BEGIN
   Id := 5;
   CancelOrders := FALSE;
   PauseOrders := FALSE;
   ResumeOrders := FALSE;
   OrderSent := FALSE;
   CurrentOrder := 0;
   NextOrder := 1;
   OrderTable[0].OrderNo := 0;
   OrderTable[0].StepNo := 256;
   OrderTable[0].PlaceTime := '';
   OrderTable[0].Device := '';
   OrderTable[0].Sequence := 0;
   OrderTable[0].Status := 'Error';
   OrderTable[0].CompleteTime := '06/10/2022 08:58:15';
   OrderTable[0].ErrorID := 0;
   OrderTable[1].OrderNo := 0;
   OrderTable[1].StepNo := 0;
   OrderTable[1].PlaceTime := '';
   OrderTable[1].Device := '';
   OrderTable[1].Sequence := 0;
   OrderTable[1].Status := '';
   OrderTable[1].CompleteTime := '';
   OrderTable[1].ErrorID := 0;
   OrderTable[2].OrderNo := 0;
   OrderTable[2].StepNo := 0;
   OrderTable[2].PlaceTime := '';
   OrderTable[2].Device := '';
   OrderTable[2].Sequence := 0;
   OrderTable[2].Status := '';
   OrderTable[2].CompleteTime := '';
   OrderTable[2].ErrorID := 0;
   OrderTable[3].OrderNo := 0;
   OrderTable[3].StepNo := 0;
   OrderTable[3].PlaceTime := '';
   OrderTable[3].Device := '';
   OrderTable[3].Sequence := 0;
   OrderTable[3].Status := '';
   OrderTable[3].CompleteTime := '';
   OrderTable[3].ErrorID := 0;
   OrderTable[4].OrderNo := 0;
   OrderTable[4].StepNo := 0;
   OrderTable[4].PlaceTime := '';
   OrderTable[4].Device := '';
   OrderTable[4].Sequence := 0;
   OrderTable[4].Status := '';
   OrderTable[4].CompleteTime := '';
   OrderTable[4].ErrorID := 0;
   OrderTable[5].OrderNo := 0;
   OrderTable[5].StepNo := 0;
   OrderTable[5].PlaceTime := '';
   OrderTable[5].Device := '';
   OrderTable[5].Sequence := 0;
   OrderTable[5].Status := '';
   OrderTable[5].CompleteTime := '';
   OrderTable[5].ErrorID := 0;
   OrderTable[6].OrderNo := 0;
   OrderTable[6].StepNo := 0;
   OrderTable[6].PlaceTime := '';
   OrderTable[6].Device := '';
   OrderTable[6].Sequence := 0;
   OrderTable[6].Status := '';
   OrderTable[6].CompleteTime := '';
   OrderTable[6].ErrorID := 0;
   OrderTable[7].OrderNo := 0;
   OrderTable[7].StepNo := 0;
   OrderTable[7].PlaceTime := '';
   OrderTable[7].Device := '';
   OrderTable[7].Sequence := 0;
   OrderTable[7].Status := '';
   OrderTable[7].CompleteTime := '';
   OrderTable[7].ErrorID := 0;
   OrderTable[8].OrderNo := 0;
   OrderTable[8].StepNo := 0;
   OrderTable[8].PlaceTime := '';
   OrderTable[8].Device := '';
   OrderTable[8].Sequence := 0;
   OrderTable[8].Status := '';
   OrderTable[8].CompleteTime := '';
   OrderTable[8].ErrorID := 0;
   OrderTable[9].OrderNo := 0;
   OrderTable[9].StepNo := 0;
   OrderTable[9].PlaceTime := '';
   OrderTable[9].Device := '';
   OrderTable[9].Sequence := 0;
   OrderTable[9].Status := '';
   OrderTable[9].CompleteTime := '';
   OrderTable[9].ErrorID := 0;
   OrderTable[10].OrderNo := 0;
   OrderTable[10].StepNo := 0;
   OrderTable[10].PlaceTime := '';
   OrderTable[10].Device := '';
   OrderTable[10].Sequence := 0;
   OrderTable[10].Status := '';
   OrderTable[10].CompleteTime := '';
   OrderTable[10].ErrorID := 0;
   OrderTable[11].OrderNo := 0;
   OrderTable[11].StepNo := 0;
   OrderTable[11].PlaceTime := '';
   OrderTable[11].Device := '';
   OrderTable[11].Sequence := 0;
   OrderTable[11].Status := '';
   OrderTable[11].CompleteTime := '';
   OrderTable[11].ErrorID := 0;
   OrderTable[12].OrderNo := 0;
   OrderTable[12].StepNo := 0;
   OrderTable[12].PlaceTime := '';
   OrderTable[12].Device := '';
   OrderTable[12].Sequence := 0;
   OrderTable[12].Status := '';
   OrderTable[12].CompleteTime := '';
   OrderTable[12].ErrorID := 0;
   OrderTable[13].OrderNo := 0;
   OrderTable[13].StepNo := 0;
   OrderTable[13].PlaceTime := '';
   OrderTable[13].Device := '';
   OrderTable[13].Sequence := 0;
   OrderTable[13].Status := '';
   OrderTable[13].CompleteTime := '';
   OrderTable[13].ErrorID := 0;
   OrderTable[14].OrderNo := 0;
   OrderTable[14].StepNo := 0;
   OrderTable[14].PlaceTime := '';
   OrderTable[14].Device := '';
   OrderTable[14].Sequence := 0;
   OrderTable[14].Status := '';
   OrderTable[14].CompleteTime := '';
   OrderTable[14].ErrorID := 0;
   OrderTable[15].OrderNo := 0;
   OrderTable[15].StepNo := 0;
   OrderTable[15].PlaceTime := '';
   OrderTable[15].Device := '';
   OrderTable[15].Sequence := 0;
   OrderTable[15].Status := '';
   OrderTable[15].CompleteTime := '';
   OrderTable[15].ErrorID := 0;
   OrderTable[16].OrderNo := 0;
   OrderTable[16].StepNo := 0;
   OrderTable[16].PlaceTime := '';
   OrderTable[16].Device := '';
   OrderTable[16].Sequence := 0;
   OrderTable[16].Status := '';
   OrderTable[16].CompleteTime := '';
   OrderTable[16].ErrorID := 0;
   OrderTable[17].OrderNo := 0;
   OrderTable[17].StepNo := 0;
   OrderTable[17].PlaceTime := '';
   OrderTable[17].Device := '';
   OrderTable[17].Sequence := 0;
   OrderTable[17].Status := '';
   OrderTable[17].CompleteTime := '';
   OrderTable[17].ErrorID := 0;
   OrderTable[18].OrderNo := 0;
   OrderTable[18].StepNo := 0;
   OrderTable[18].PlaceTime := '';
   OrderTable[18].Device := '';
   OrderTable[18].Sequence := 0;
   OrderTable[18].Status := '';
   OrderTable[18].CompleteTime := '';
   OrderTable[18].ErrorID := 0;
   OrderTable[19].OrderNo := 0;
   OrderTable[19].StepNo := 0;
   OrderTable[19].PlaceTime := '';
   OrderTable[19].Device := '';
   OrderTable[19].Sequence := 0;
   OrderTable[19].Status := '';
   OrderTable[19].CompleteTime := '';
   OrderTable[19].ErrorID := 0;
   OrderTable[20].OrderNo := 0;
   OrderTable[20].StepNo := 0;
   OrderTable[20].PlaceTime := '';
   OrderTable[20].Device := '';
   OrderTable[20].Sequence := 0;
   OrderTable[20].Status := '';
   OrderTable[20].CompleteTime := '';
   OrderTable[20].ErrorID := 0;
   OrderTable[21].OrderNo := 0;
   OrderTable[21].StepNo := 0;
   OrderTable[21].PlaceTime := '';
   OrderTable[21].Device := '';
   OrderTable[21].Sequence := 0;
   OrderTable[21].Status := '';
   OrderTable[21].CompleteTime := '';
   OrderTable[21].ErrorID := 0;
   OrderTable[22].OrderNo := 0;
   OrderTable[22].StepNo := 0;
   OrderTable[22].PlaceTime := '';
   OrderTable[22].Device := '';
   OrderTable[22].Sequence := 0;
   OrderTable[22].Status := '';
   OrderTable[22].CompleteTime := '';
   OrderTable[22].ErrorID := 0;
   OrderTable[23].OrderNo := 0;
   OrderTable[23].StepNo := 0;
   OrderTable[23].PlaceTime := '';
   OrderTable[23].Device := '';
   OrderTable[23].Sequence := 0;
   OrderTable[23].Status := '';
   OrderTable[23].CompleteTime := '';
   OrderTable[23].ErrorID := 0;
   OrderTable[24].OrderNo := 0;
   OrderTable[24].StepNo := 0;
   OrderTable[24].PlaceTime := '';
   OrderTable[24].Device := '';
   OrderTable[24].Sequence := 0;
   OrderTable[24].Status := '';
   OrderTable[24].CompleteTime := '';
   OrderTable[24].ErrorID := 0;
   OrderTable[25].OrderNo := 0;
   OrderTable[25].StepNo := 0;
   OrderTable[25].PlaceTime := '';
   OrderTable[25].Device := '';
   OrderTable[25].Sequence := 0;
   OrderTable[25].Status := '';
   OrderTable[25].CompleteTime := '';
   OrderTable[25].ErrorID := 0;
   OrderTable[26].OrderNo := 0;
   OrderTable[26].StepNo := 0;
   OrderTable[26].PlaceTime := '';
   OrderTable[26].Device := '';
   OrderTable[26].Sequence := 0;
   OrderTable[26].Status := '';
   OrderTable[26].CompleteTime := '';
   OrderTable[26].ErrorID := 0;
   OrderTable[27].OrderNo := 0;
   OrderTable[27].StepNo := 0;
   OrderTable[27].PlaceTime := '';
   OrderTable[27].Device := '';
   OrderTable[27].Sequence := 0;
   OrderTable[27].Status := '';
   OrderTable[27].CompleteTime := '';
   OrderTable[27].ErrorID := 0;
   OrderTable[28].OrderNo := 0;
   OrderTable[28].StepNo := 0;
   OrderTable[28].PlaceTime := '';
   OrderTable[28].Device := '';
   OrderTable[28].Sequence := 0;
   OrderTable[28].Status := '';
   OrderTable[28].CompleteTime := '';
   OrderTable[28].ErrorID := 0;
   OrderTable[29].OrderNo := 0;
   OrderTable[29].StepNo := 0;
   OrderTable[29].PlaceTime := '';
   OrderTable[29].Device := '';
   OrderTable[29].Sequence := 0;
   OrderTable[29].Status := '';
   OrderTable[29].CompleteTime := '';
   OrderTable[29].ErrorID := 0;
   OrderTable[30].OrderNo := 0;
   OrderTable[30].StepNo := 0;
   OrderTable[30].PlaceTime := '';
   OrderTable[30].Device := '';
   OrderTable[30].Sequence := 0;
   OrderTable[30].Status := '';
   OrderTable[30].CompleteTime := '';
   OrderTable[30].ErrorID := 0;
   OrderTable[31].OrderNo := 0;
   OrderTable[31].StepNo := 0;
   OrderTable[31].PlaceTime := '';
   OrderTable[31].Device := '';
   OrderTable[31].Sequence := 0;
   OrderTable[31].Status := '';
   OrderTable[31].CompleteTime := '';
   OrderTable[31].ErrorID := 0;
   OrderTable[32].OrderNo := 0;
   OrderTable[32].StepNo := 0;
   OrderTable[32].PlaceTime := '';
   OrderTable[32].Device := '';
   OrderTable[32].Sequence := 0;
   OrderTable[32].Status := '';
   OrderTable[32].CompleteTime := '';
   OrderTable[32].ErrorID := 0;
   OrderTable[33].OrderNo := 0;
   OrderTable[33].StepNo := 0;
   OrderTable[33].PlaceTime := '';
   OrderTable[33].Device := '';
   OrderTable[33].Sequence := 0;
   OrderTable[33].Status := '';
   OrderTable[33].CompleteTime := '';
   OrderTable[33].ErrorID := 0;
   OrderTable[34].OrderNo := 0;
   OrderTable[34].StepNo := 0;
   OrderTable[34].PlaceTime := '';
   OrderTable[34].Device := '';
   OrderTable[34].Sequence := 0;
   OrderTable[34].Status := '';
   OrderTable[34].CompleteTime := '';
   OrderTable[34].ErrorID := 0;
   OrderTable[35].OrderNo := 0;
   OrderTable[35].StepNo := 0;
   OrderTable[35].PlaceTime := '';
   OrderTable[35].Device := '';
   OrderTable[35].Sequence := 0;
   OrderTable[35].Status := '';
   OrderTable[35].CompleteTime := '';
   OrderTable[35].ErrorID := 0;
   OrderTable[36].OrderNo := 0;
   OrderTable[36].StepNo := 0;
   OrderTable[36].PlaceTime := '';
   OrderTable[36].Device := '';
   OrderTable[36].Sequence := 0;
   OrderTable[36].Status := '';
   OrderTable[36].CompleteTime := '';
   OrderTable[36].ErrorID := 0;
   OrderTable[37].OrderNo := 0;
   OrderTable[37].StepNo := 0;
   OrderTable[37].PlaceTime := '';
   OrderTable[37].Device := '';
   OrderTable[37].Sequence := 0;
   OrderTable[37].Status := '';
   OrderTable[37].CompleteTime := '';
   OrderTable[37].ErrorID := 0;
   OrderTable[38].OrderNo := 0;
   OrderTable[38].StepNo := 0;
   OrderTable[38].PlaceTime := '';
   OrderTable[38].Device := '';
   OrderTable[38].Sequence := 0;
   OrderTable[38].Status := '';
   OrderTable[38].CompleteTime := '';
   OrderTable[38].ErrorID := 0;
   OrderTable[39].OrderNo := 0;
   OrderTable[39].StepNo := 0;
   OrderTable[39].PlaceTime := '';
   OrderTable[39].Device := '';
   OrderTable[39].Sequence := 0;
   OrderTable[39].Status := '';
   OrderTable[39].CompleteTime := '';
   OrderTable[39].ErrorID := 0;
   OrderTable[40].OrderNo := 0;
   OrderTable[40].StepNo := 0;
   OrderTable[40].PlaceTime := '';
   OrderTable[40].Device := '';
   OrderTable[40].Sequence := 0;
   OrderTable[40].Status := '';
   OrderTable[40].CompleteTime := '';
   OrderTable[40].ErrorID := 0;
   OrderTable[41].OrderNo := 0;
   OrderTable[41].StepNo := 0;
   OrderTable[41].PlaceTime := '';
   OrderTable[41].Device := '';
   OrderTable[41].Sequence := 0;
   OrderTable[41].Status := '';
   OrderTable[41].CompleteTime := '';
   OrderTable[41].ErrorID := 0;
   OrderTable[42].OrderNo := 0;
   OrderTable[42].StepNo := 0;
   OrderTable[42].PlaceTime := '';
   OrderTable[42].Device := '';
   OrderTable[42].Sequence := 0;
   OrderTable[42].Status := '';
   OrderTable[42].CompleteTime := '';
   OrderTable[42].ErrorID := 0;
   OrderTable[43].OrderNo := 0;
   OrderTable[43].StepNo := 0;
   OrderTable[43].PlaceTime := '';
   OrderTable[43].Device := '';
   OrderTable[43].Sequence := 0;
   OrderTable[43].Status := '';
   OrderTable[43].CompleteTime := '';
   OrderTable[43].ErrorID := 0;
   OrderTable[44].OrderNo := 0;
   OrderTable[44].StepNo := 0;
   OrderTable[44].PlaceTime := '';
   OrderTable[44].Device := '';
   OrderTable[44].Sequence := 0;
   OrderTable[44].Status := '';
   OrderTable[44].CompleteTime := '';
   OrderTable[44].ErrorID := 0;
   OrderTable[45].OrderNo := 0;
   OrderTable[45].StepNo := 0;
   OrderTable[45].PlaceTime := '';
   OrderTable[45].Device := '';
   OrderTable[45].Sequence := 0;
   OrderTable[45].Status := '';
   OrderTable[45].CompleteTime := '';
   OrderTable[45].ErrorID := 0;
   OrderTable[46].OrderNo := 0;
   OrderTable[46].StepNo := 0;
   OrderTable[46].PlaceTime := '';
   OrderTable[46].Device := '';
   OrderTable[46].Sequence := 0;
   OrderTable[46].Status := '';
   OrderTable[46].CompleteTime := '';
   OrderTable[46].ErrorID := 0;
   OrderTable[47].OrderNo := 0;
   OrderTable[47].StepNo := 0;
   OrderTable[47].PlaceTime := '';
   OrderTable[47].Device := '';
   OrderTable[47].Sequence := 0;
   OrderTable[47].Status := '';
   OrderTable[47].CompleteTime := '';
   OrderTable[47].ErrorID := 0;
   OrderTable[48].OrderNo := 0;
   OrderTable[48].StepNo := 0;
   OrderTable[48].PlaceTime := '';
   OrderTable[48].Device := '';
   OrderTable[48].Sequence := 0;
   OrderTable[48].Status := '';
   OrderTable[48].CompleteTime := '';
   OrderTable[48].ErrorID := 0;
   OrderTable[49].OrderNo := 0;
   OrderTable[49].StepNo := 0;
   OrderTable[49].PlaceTime := '';
   OrderTable[49].Device := '';
   OrderTable[49].Sequence := 0;
   OrderTable[49].Status := '';
   OrderTable[49].CompleteTime := '';
   OrderTable[49].ErrorID := 0;
   OrderTable[50].OrderNo := 0;
   OrderTable[50].StepNo := 0;
   OrderTable[50].PlaceTime := '';
   OrderTable[50].Device := '';
   OrderTable[50].Sequence := 0;
   OrderTable[50].Status := '';
   OrderTable[50].CompleteTime := '';
   OrderTable[50].ErrorID := 0;
   OrderTable[51].OrderNo := 0;
   OrderTable[51].StepNo := 0;
   OrderTable[51].PlaceTime := '';
   OrderTable[51].Device := '';
   OrderTable[51].Sequence := 0;
   OrderTable[51].Status := '';
   OrderTable[51].CompleteTime := '';
   OrderTable[51].ErrorID := 0;
   OrderTable[52].OrderNo := 0;
   OrderTable[52].StepNo := 0;
   OrderTable[52].PlaceTime := '';
   OrderTable[52].Device := '';
   OrderTable[52].Sequence := 0;
   OrderTable[52].Status := '';
   OrderTable[52].CompleteTime := '';
   OrderTable[52].ErrorID := 0;
   OrderTable[53].OrderNo := 0;
   OrderTable[53].StepNo := 0;
   OrderTable[53].PlaceTime := '';
   OrderTable[53].Device := '';
   OrderTable[53].Sequence := 0;
   OrderTable[53].Status := '';
   OrderTable[53].CompleteTime := '';
   OrderTable[53].ErrorID := 0;
   OrderTable[54].OrderNo := 0;
   OrderTable[54].StepNo := 0;
   OrderTable[54].PlaceTime := '';
   OrderTable[54].Device := '';
   OrderTable[54].Sequence := 0;
   OrderTable[54].Status := '';
   OrderTable[54].CompleteTime := '';
   OrderTable[54].ErrorID := 0;
   OrderTable[55].OrderNo := 0;
   OrderTable[55].StepNo := 0;
   OrderTable[55].PlaceTime := '';
   OrderTable[55].Device := '';
   OrderTable[55].Sequence := 0;
   OrderTable[55].Status := '';
   OrderTable[55].CompleteTime := '';
   OrderTable[55].ErrorID := 0;
   OrderTable[56].OrderNo := 0;
   OrderTable[56].StepNo := 0;
   OrderTable[56].PlaceTime := '';
   OrderTable[56].Device := '';
   OrderTable[56].Sequence := 0;
   OrderTable[56].Status := '';
   OrderTable[56].CompleteTime := '';
   OrderTable[56].ErrorID := 0;
   OrderTable[57].OrderNo := 0;
   OrderTable[57].StepNo := 0;
   OrderTable[57].PlaceTime := '';
   OrderTable[57].Device := '';
   OrderTable[57].Sequence := 0;
   OrderTable[57].Status := '';
   OrderTable[57].CompleteTime := '';
   OrderTable[57].ErrorID := 0;
   OrderTable[58].OrderNo := 0;
   OrderTable[58].StepNo := 0;
   OrderTable[58].PlaceTime := '';
   OrderTable[58].Device := '';
   OrderTable[58].Sequence := 0;
   OrderTable[58].Status := '';
   OrderTable[58].CompleteTime := '';
   OrderTable[58].ErrorID := 0;
   OrderTable[59].OrderNo := 0;
   OrderTable[59].StepNo := 0;
   OrderTable[59].PlaceTime := '';
   OrderTable[59].Device := '';
   OrderTable[59].Sequence := 0;
   OrderTable[59].Status := '';
   OrderTable[59].CompleteTime := '';
   OrderTable[59].ErrorID := 0;
   OrderTable[60].OrderNo := 0;
   OrderTable[60].StepNo := 0;
   OrderTable[60].PlaceTime := '';
   OrderTable[60].Device := '';
   OrderTable[60].Sequence := 0;
   OrderTable[60].Status := '';
   OrderTable[60].CompleteTime := '';
   OrderTable[60].ErrorID := 0;
   OrderTable[61].OrderNo := 0;
   OrderTable[61].StepNo := 0;
   OrderTable[61].PlaceTime := '';
   OrderTable[61].Device := '';
   OrderTable[61].Sequence := 0;
   OrderTable[61].Status := '';
   OrderTable[61].CompleteTime := '';
   OrderTable[61].ErrorID := 0;
   OrderTable[62].OrderNo := 0;
   OrderTable[62].StepNo := 0;
   OrderTable[62].PlaceTime := '';
   OrderTable[62].Device := '';
   OrderTable[62].Sequence := 0;
   OrderTable[62].Status := '';
   OrderTable[62].CompleteTime := '';
   OrderTable[62].ErrorID := 0;
   OrderTable[63].OrderNo := 0;
   OrderTable[63].StepNo := 0;
   OrderTable[63].PlaceTime := '';
   OrderTable[63].Device := '';
   OrderTable[63].Sequence := 0;
   OrderTable[63].Status := '';
   OrderTable[63].CompleteTime := '';
   OrderTable[63].ErrorID := 0;
   OrderTable[64].OrderNo := 0;
   OrderTable[64].StepNo := 0;
   OrderTable[64].PlaceTime := '';
   OrderTable[64].Device := '';
   OrderTable[64].Sequence := 0;
   OrderTable[64].Status := '';
   OrderTable[64].CompleteTime := '';
   OrderTable[64].ErrorID := 0;
   OrderTable[65].OrderNo := 0;
   OrderTable[65].StepNo := 0;
   OrderTable[65].PlaceTime := '';
   OrderTable[65].Device := '';
   OrderTable[65].Sequence := 0;
   OrderTable[65].Status := '';
   OrderTable[65].CompleteTime := '';
   OrderTable[65].ErrorID := 0;
   OrderTable[66].OrderNo := 0;
   OrderTable[66].StepNo := 0;
   OrderTable[66].PlaceTime := '';
   OrderTable[66].Device := '';
   OrderTable[66].Sequence := 0;
   OrderTable[66].Status := '';
   OrderTable[66].CompleteTime := '';
   OrderTable[66].ErrorID := 0;
   OrderTable[67].OrderNo := 0;
   OrderTable[67].StepNo := 0;
   OrderTable[67].PlaceTime := '';
   OrderTable[67].Device := '';
   OrderTable[67].Sequence := 0;
   OrderTable[67].Status := '';
   OrderTable[67].CompleteTime := '';
   OrderTable[67].ErrorID := 0;
   OrderTable[68].OrderNo := 0;
   OrderTable[68].StepNo := 0;
   OrderTable[68].PlaceTime := '';
   OrderTable[68].Device := '';
   OrderTable[68].Sequence := 0;
   OrderTable[68].Status := '';
   OrderTable[68].CompleteTime := '';
   OrderTable[68].ErrorID := 0;
   OrderTable[69].OrderNo := 0;
   OrderTable[69].StepNo := 0;
   OrderTable[69].PlaceTime := '';
   OrderTable[69].Device := '';
   OrderTable[69].Sequence := 0;
   OrderTable[69].Status := '';
   OrderTable[69].CompleteTime := '';
   OrderTable[69].ErrorID := 0;
   OrderTable[70].OrderNo := 0;
   OrderTable[70].StepNo := 0;
   OrderTable[70].PlaceTime := '';
   OrderTable[70].Device := '';
   OrderTable[70].Sequence := 0;
   OrderTable[70].Status := '';
   OrderTable[70].CompleteTime := '';
   OrderTable[70].ErrorID := 0;
   OrderTable[71].OrderNo := 0;
   OrderTable[71].StepNo := 0;
   OrderTable[71].PlaceTime := '';
   OrderTable[71].Device := '';
   OrderTable[71].Sequence := 0;
   OrderTable[71].Status := '';
   OrderTable[71].CompleteTime := '';
   OrderTable[71].ErrorID := 0;
   OrderTable[72].OrderNo := 0;
   OrderTable[72].StepNo := 0;
   OrderTable[72].PlaceTime := '';
   OrderTable[72].Device := '';
   OrderTable[72].Sequence := 0;
   OrderTable[72].Status := '';
   OrderTable[72].CompleteTime := '';
   OrderTable[72].ErrorID := 0;
   OrderTable[73].OrderNo := 0;
   OrderTable[73].StepNo := 0;
   OrderTable[73].PlaceTime := '';
   OrderTable[73].Device := '';
   OrderTable[73].Sequence := 0;
   OrderTable[73].Status := '';
   OrderTable[73].CompleteTime := '';
   OrderTable[73].ErrorID := 0;
   OrderTable[74].OrderNo := 0;
   OrderTable[74].StepNo := 0;
   OrderTable[74].PlaceTime := '';
   OrderTable[74].Device := '';
   OrderTable[74].Sequence := 0;
   OrderTable[74].Status := '';
   OrderTable[74].CompleteTime := '';
   OrderTable[74].ErrorID := 0;
   OrderTable[75].OrderNo := 0;
   OrderTable[75].StepNo := 0;
   OrderTable[75].PlaceTime := '';
   OrderTable[75].Device := '';
   OrderTable[75].Sequence := 0;
   OrderTable[75].Status := '';
   OrderTable[75].CompleteTime := '';
   OrderTable[75].ErrorID := 0;
   OrderTable[76].OrderNo := 0;
   OrderTable[76].StepNo := 0;
   OrderTable[76].PlaceTime := '';
   OrderTable[76].Device := '';
   OrderTable[76].Sequence := 0;
   OrderTable[76].Status := '';
   OrderTable[76].CompleteTime := '';
   OrderTable[76].ErrorID := 0;
   OrderTable[77].OrderNo := 0;
   OrderTable[77].StepNo := 0;
   OrderTable[77].PlaceTime := '';
   OrderTable[77].Device := '';
   OrderTable[77].Sequence := 0;
   OrderTable[77].Status := '';
   OrderTable[77].CompleteTime := '';
   OrderTable[77].ErrorID := 0;
   OrderTable[78].OrderNo := 0;
   OrderTable[78].StepNo := 0;
   OrderTable[78].PlaceTime := '';
   OrderTable[78].Device := '';
   OrderTable[78].Sequence := 0;
   OrderTable[78].Status := '';
   OrderTable[78].CompleteTime := '';
   OrderTable[78].ErrorID := 0;
   OrderTable[79].OrderNo := 0;
   OrderTable[79].StepNo := 0;
   OrderTable[79].PlaceTime := '';
   OrderTable[79].Device := '';
   OrderTable[79].Sequence := 0;
   OrderTable[79].Status := '';
   OrderTable[79].CompleteTime := '';
   OrderTable[79].ErrorID := 0;
   OrderTable[80].OrderNo := 0;
   OrderTable[80].StepNo := 0;
   OrderTable[80].PlaceTime := '';
   OrderTable[80].Device := '';
   OrderTable[80].Sequence := 0;
   OrderTable[80].Status := '';
   OrderTable[80].CompleteTime := '';
   OrderTable[80].ErrorID := 0;
   OrderTable[81].OrderNo := 0;
   OrderTable[81].StepNo := 0;
   OrderTable[81].PlaceTime := '';
   OrderTable[81].Device := '';
   OrderTable[81].Sequence := 0;
   OrderTable[81].Status := '';
   OrderTable[81].CompleteTime := '';
   OrderTable[81].ErrorID := 0;
   OrderTable[82].OrderNo := 0;
   OrderTable[82].StepNo := 0;
   OrderTable[82].PlaceTime := '';
   OrderTable[82].Device := '';
   OrderTable[82].Sequence := 0;
   OrderTable[82].Status := '';
   OrderTable[82].CompleteTime := '';
   OrderTable[82].ErrorID := 0;
   OrderTable[83].OrderNo := 0;
   OrderTable[83].StepNo := 0;
   OrderTable[83].PlaceTime := '';
   OrderTable[83].Device := '';
   OrderTable[83].Sequence := 0;
   OrderTable[83].Status := '';
   OrderTable[83].CompleteTime := '';
   OrderTable[83].ErrorID := 0;
   OrderTable[84].OrderNo := 0;
   OrderTable[84].StepNo := 0;
   OrderTable[84].PlaceTime := '';
   OrderTable[84].Device := '';
   OrderTable[84].Sequence := 0;
   OrderTable[84].Status := '';
   OrderTable[84].CompleteTime := '';
   OrderTable[84].ErrorID := 0;
   OrderTable[85].OrderNo := 0;
   OrderTable[85].StepNo := 0;
   OrderTable[85].PlaceTime := '';
   OrderTable[85].Device := '';
   OrderTable[85].Sequence := 0;
   OrderTable[85].Status := '';
   OrderTable[85].CompleteTime := '';
   OrderTable[85].ErrorID := 0;
   OrderTable[86].OrderNo := 0;
   OrderTable[86].StepNo := 0;
   OrderTable[86].PlaceTime := '';
   OrderTable[86].Device := '';
   OrderTable[86].Sequence := 0;
   OrderTable[86].Status := '';
   OrderTable[86].CompleteTime := '';
   OrderTable[86].ErrorID := 0;
   OrderTable[87].OrderNo := 0;
   OrderTable[87].StepNo := 0;
   OrderTable[87].PlaceTime := '';
   OrderTable[87].Device := '';
   OrderTable[87].Sequence := 0;
   OrderTable[87].Status := '';
   OrderTable[87].CompleteTime := '';
   OrderTable[87].ErrorID := 0;
   OrderTable[88].OrderNo := 0;
   OrderTable[88].StepNo := 0;
   OrderTable[88].PlaceTime := '';
   OrderTable[88].Device := '';
   OrderTable[88].Sequence := 0;
   OrderTable[88].Status := '';
   OrderTable[88].CompleteTime := '';
   OrderTable[88].ErrorID := 0;
   OrderTable[89].OrderNo := 0;
   OrderTable[89].StepNo := 0;
   OrderTable[89].PlaceTime := '';
   OrderTable[89].Device := '';
   OrderTable[89].Sequence := 0;
   OrderTable[89].Status := '';
   OrderTable[89].CompleteTime := '';
   OrderTable[89].ErrorID := 0;
   OrderTable[90].OrderNo := 0;
   OrderTable[90].StepNo := 0;
   OrderTable[90].PlaceTime := '';
   OrderTable[90].Device := '';
   OrderTable[90].Sequence := 0;
   OrderTable[90].Status := '';
   OrderTable[90].CompleteTime := '';
   OrderTable[90].ErrorID := 0;
   OrderTable[91].OrderNo := 0;
   OrderTable[91].StepNo := 0;
   OrderTable[91].PlaceTime := '';
   OrderTable[91].Device := '';
   OrderTable[91].Sequence := 0;
   OrderTable[91].Status := '';
   OrderTable[91].CompleteTime := '';
   OrderTable[91].ErrorID := 0;
   OrderTable[92].OrderNo := 0;
   OrderTable[92].StepNo := 0;
   OrderTable[92].PlaceTime := '';
   OrderTable[92].Device := '';
   OrderTable[92].Sequence := 0;
   OrderTable[92].Status := '';
   OrderTable[92].CompleteTime := '';
   OrderTable[92].ErrorID := 0;
   OrderTable[93].OrderNo := 0;
   OrderTable[93].StepNo := 0;
   OrderTable[93].PlaceTime := '';
   OrderTable[93].Device := '';
   OrderTable[93].Sequence := 0;
   OrderTable[93].Status := '';
   OrderTable[93].CompleteTime := '';
   OrderTable[93].ErrorID := 0;
   OrderTable[94].OrderNo := 0;
   OrderTable[94].StepNo := 0;
   OrderTable[94].PlaceTime := '';
   OrderTable[94].Device := '';
   OrderTable[94].Sequence := 0;
   OrderTable[94].Status := '';
   OrderTable[94].CompleteTime := '';
   OrderTable[94].ErrorID := 0;
   OrderTable[95].OrderNo := 0;
   OrderTable[95].StepNo := 0;
   OrderTable[95].PlaceTime := '';
   OrderTable[95].Device := '';
   OrderTable[95].Sequence := 0;
   OrderTable[95].Status := '';
   OrderTable[95].CompleteTime := '';
   OrderTable[95].ErrorID := 0;
   OrderTable[96].OrderNo := 0;
   OrderTable[96].StepNo := 0;
   OrderTable[96].PlaceTime := '';
   OrderTable[96].Device := '';
   OrderTable[96].Sequence := 0;
   OrderTable[96].Status := '';
   OrderTable[96].CompleteTime := '';
   OrderTable[96].ErrorID := 0;
   OrderTable[97].OrderNo := 0;
   OrderTable[97].StepNo := 0;
   OrderTable[97].PlaceTime := '';
   OrderTable[97].Device := '';
   OrderTable[97].Sequence := 0;
   OrderTable[97].Status := '';
   OrderTable[97].CompleteTime := '';
   OrderTable[97].ErrorID := 0;
   OrderTable[98].OrderNo := 0;
   OrderTable[98].StepNo := 0;
   OrderTable[98].PlaceTime := '';
   OrderTable[98].Device := '';
   OrderTable[98].Sequence := 0;
   OrderTable[98].Status := '';
   OrderTable[98].CompleteTime := '';
   OrderTable[98].ErrorID := 0;
   OrderTable[99].OrderNo := 0;
   OrderTable[99].StepNo := 0;
   OrderTable[99].PlaceTime := '';
   OrderTable[99].Device := '';
   OrderTable[99].Sequence := 0;
   OrderTable[99].Status := '';
   OrderTable[99].CompleteTime := '';
   OrderTable[99].ErrorID := 0;
   StepTable[1].OrderNo := 0;
   StepTable[1].StepNo := 0;
   StepTable[1].PlaceTime := '';
   StepTable[1].Device := '';
   StepTable[1].Sequence := 0;
   StepTable[1].Status := '';
   StepTable[1].CompleteTime := '';
   StepTable[1].ErrorID := 0;
   StepTable[2].OrderNo := 0;
   StepTable[2].StepNo := 0;
   StepTable[2].PlaceTime := '';
   StepTable[2].Device := '';
   StepTable[2].Sequence := 0;
   StepTable[2].Status := '';
   StepTable[2].CompleteTime := '';
   StepTable[2].ErrorID := 0;
   StepTable[3].OrderNo := 0;
   StepTable[3].StepNo := 0;
   StepTable[3].PlaceTime := '';
   StepTable[3].Device := '';
   StepTable[3].Sequence := 0;
   StepTable[3].Status := '';
   StepTable[3].CompleteTime := '';
   StepTable[3].ErrorID := 0;
   StepTable[4].OrderNo := 0;
   StepTable[4].StepNo := 0;
   StepTable[4].PlaceTime := '';
   StepTable[4].Device := '';
   StepTable[4].Sequence := 0;
   StepTable[4].Status := '';
   StepTable[4].CompleteTime := '';
   StepTable[4].ErrorID := 0;
   StepTable[5].OrderNo := 0;
   StepTable[5].StepNo := 0;
   StepTable[5].PlaceTime := '';
   StepTable[5].Device := '';
   StepTable[5].Sequence := 0;
   StepTable[5].Status := '';
   StepTable[5].CompleteTime := '';
   StepTable[5].ErrorID := 0;
   StepTable[6].OrderNo := 0;
   StepTable[6].StepNo := 0;
   StepTable[6].PlaceTime := '';
   StepTable[6].Device := '';
   StepTable[6].Sequence := 0;
   StepTable[6].Status := '';
   StepTable[6].CompleteTime := '';
   StepTable[6].ErrorID := 0;
   StepTable[7].OrderNo := 0;
   StepTable[7].StepNo := 0;
   StepTable[7].PlaceTime := '';
   StepTable[7].Device := '';
   StepTable[7].Sequence := 0;
   StepTable[7].Status := '';
   StepTable[7].CompleteTime := '';
   StepTable[7].ErrorID := 0;
   StepTable[8].OrderNo := 0;
   StepTable[8].StepNo := 0;
   StepTable[8].PlaceTime := '';
   StepTable[8].Device := '';
   StepTable[8].Sequence := 0;
   StepTable[8].Status := '';
   StepTable[8].CompleteTime := '';
   StepTable[8].ErrorID := 0;
   StepTable[9].OrderNo := 0;
   StepTable[9].StepNo := 0;
   StepTable[9].PlaceTime := '';
   StepTable[9].Device := '';
   StepTable[9].Sequence := 0;
   StepTable[9].Status := '';
   StepTable[9].CompleteTime := '';
   StepTable[9].ErrorID := 0;
   StepTable[10].OrderNo := 0;
   StepTable[10].StepNo := 0;
   StepTable[10].PlaceTime := '';
   StepTable[10].Device := '';
   StepTable[10].Sequence := 0;
   StepTable[10].Status := '';
   StepTable[10].CompleteTime := '';
   StepTable[10].ErrorID := 0;
   StepTable[11].OrderNo := 0;
   StepTable[11].StepNo := 0;
   StepTable[11].PlaceTime := '';
   StepTable[11].Device := '';
   StepTable[11].Sequence := 0;
   StepTable[11].Status := '';
   StepTable[11].CompleteTime := '';
   StepTable[11].ErrorID := 0;
   StepTable[12].OrderNo := 0;
   StepTable[12].StepNo := 0;
   StepTable[12].PlaceTime := '';
   StepTable[12].Device := '';
   StepTable[12].Sequence := 0;
   StepTable[12].Status := '';
   StepTable[12].CompleteTime := '';
   StepTable[12].ErrorID := 0;
   StepTable[13].OrderNo := 0;
   StepTable[13].StepNo := 0;
   StepTable[13].PlaceTime := '';
   StepTable[13].Device := '';
   StepTable[13].Sequence := 0;
   StepTable[13].Status := '';
   StepTable[13].CompleteTime := '';
   StepTable[13].ErrorID := 0;
   StepTable[14].OrderNo := 0;
   StepTable[14].StepNo := 0;
   StepTable[14].PlaceTime := '';
   StepTable[14].Device := '';
   StepTable[14].Sequence := 0;
   StepTable[14].Status := '';
   StepTable[14].CompleteTime := '';
   StepTable[14].ErrorID := 0;
   StepTable[15].OrderNo := 0;
   StepTable[15].StepNo := 0;
   StepTable[15].PlaceTime := '';
   StepTable[15].Device := '';
   StepTable[15].Sequence := 0;
   StepTable[15].Status := '';
   StepTable[15].CompleteTime := '';
   StepTable[15].ErrorID := 0;
   StepTable[16].OrderNo := 0;
   StepTable[16].StepNo := 0;
   StepTable[16].PlaceTime := '';
   StepTable[16].Device := '';
   StepTable[16].Sequence := 0;
   StepTable[16].Status := '';
   StepTable[16].CompleteTime := '';
   StepTable[16].ErrorID := 0;
   StepTable[17].OrderNo := 0;
   StepTable[17].StepNo := 0;
   StepTable[17].PlaceTime := '';
   StepTable[17].Device := '';
   StepTable[17].Sequence := 0;
   StepTable[17].Status := '';
   StepTable[17].CompleteTime := '';
   StepTable[17].ErrorID := 0;
   StepTable[18].OrderNo := 0;
   StepTable[18].StepNo := 0;
   StepTable[18].PlaceTime := '';
   StepTable[18].Device := '';
   StepTable[18].Sequence := 0;
   StepTable[18].Status := '';
   StepTable[18].CompleteTime := '';
   StepTable[18].ErrorID := 0;
   StepTable[19].OrderNo := 0;
   StepTable[19].StepNo := 0;
   StepTable[19].PlaceTime := '';
   StepTable[19].Device := '';
   StepTable[19].Sequence := 0;
   StepTable[19].Status := '';
   StepTable[19].CompleteTime := '';
   StepTable[19].ErrorID := 0;
   StepTable[20].OrderNo := 0;
   StepTable[20].StepNo := 0;
   StepTable[20].PlaceTime := '';
   StepTable[20].Device := '';
   StepTable[20].Sequence := 0;
   StepTable[20].Status := '';
   StepTable[20].CompleteTime := '';
   StepTable[20].ErrorID := 0;
   CarParked_Confirm := FALSE;
   Running := FALSE;
   IDLE := TRUE;
   Error := FALSE;
   State := 0;
   ResetError := FALSE;
   Ready := TRUE;
   Selected := TRUE;
   Auto_Man := TRUE;
   Paused := FALSE;

END_DATA_BLOCK

DATA_BLOCK "Auto_Test_2_DB"
{ S7_Optimized_Access := 'TRUE' }
VERSION : 0.1
NON_RETAIN
"Auto_Test"

BEGIN

END_DATA_BLOCK

DATA_BLOCK "System_DB_4"
{ S7_Optimized_Access := 'TRUE' }
VERSION : 0.1
NON_RETAIN
"System_UDT"

BEGIN
   Id := 4;
   CancelOrders := FALSE;
   PauseOrders := FALSE;
   ResumeOrders := FALSE;
   OrderSent := FALSE;
   CurrentOrder := 0;
   NextOrder := 1;
   OrderTable[0].OrderNo := 0;
   OrderTable[0].StepNo := 256;
   OrderTable[0].PlaceTime := '';
   OrderTable[0].Device := '';
   OrderTable[0].Sequence := 0;
   OrderTable[0].Status := 'Error';
   OrderTable[0].CompleteTime := '06/10/2022 08:58:15';
   OrderTable[0].ErrorID := 0;
   OrderTable[1].OrderNo := 0;
   OrderTable[1].StepNo := 0;
   OrderTable[1].PlaceTime := '';
   OrderTable[1].Device := '';
   OrderTable[1].Sequence := 0;
   OrderTable[1].Status := '';
   OrderTable[1].CompleteTime := '';
   OrderTable[1].ErrorID := 0;
   OrderTable[2].OrderNo := 0;
   OrderTable[2].StepNo := 0;
   OrderTable[2].PlaceTime := '';
   OrderTable[2].Device := '';
   OrderTable[2].Sequence := 0;
   OrderTable[2].Status := '';
   OrderTable[2].CompleteTime := '';
   OrderTable[2].ErrorID := 0;
   OrderTable[3].OrderNo := 0;
   OrderTable[3].StepNo := 0;
   OrderTable[3].PlaceTime := '';
   OrderTable[3].Device := '';
   OrderTable[3].Sequence := 0;
   OrderTable[3].Status := '';
   OrderTable[3].CompleteTime := '';
   OrderTable[3].ErrorID := 0;
   OrderTable[4].OrderNo := 0;
   OrderTable[4].StepNo := 0;
   OrderTable[4].PlaceTime := '';
   OrderTable[4].Device := '';
   OrderTable[4].Sequence := 0;
   OrderTable[4].Status := '';
   OrderTable[4].CompleteTime := '';
   OrderTable[4].ErrorID := 0;
   OrderTable[5].OrderNo := 0;
   OrderTable[5].StepNo := 0;
   OrderTable[5].PlaceTime := '';
   OrderTable[5].Device := '';
   OrderTable[5].Sequence := 0;
   OrderTable[5].Status := '';
   OrderTable[5].CompleteTime := '';
   OrderTable[5].ErrorID := 0;
   OrderTable[6].OrderNo := 0;
   OrderTable[6].StepNo := 0;
   OrderTable[6].PlaceTime := '';
   OrderTable[6].Device := '';
   OrderTable[6].Sequence := 0;
   OrderTable[6].Status := '';
   OrderTable[6].CompleteTime := '';
   OrderTable[6].ErrorID := 0;
   OrderTable[7].OrderNo := 0;
   OrderTable[7].StepNo := 0;
   OrderTable[7].PlaceTime := '';
   OrderTable[7].Device := '';
   OrderTable[7].Sequence := 0;
   OrderTable[7].Status := '';
   OrderTable[7].CompleteTime := '';
   OrderTable[7].ErrorID := 0;
   OrderTable[8].OrderNo := 0;
   OrderTable[8].StepNo := 0;
   OrderTable[8].PlaceTime := '';
   OrderTable[8].Device := '';
   OrderTable[8].Sequence := 0;
   OrderTable[8].Status := '';
   OrderTable[8].CompleteTime := '';
   OrderTable[8].ErrorID := 0;
   OrderTable[9].OrderNo := 0;
   OrderTable[9].StepNo := 0;
   OrderTable[9].PlaceTime := '';
   OrderTable[9].Device := '';
   OrderTable[9].Sequence := 0;
   OrderTable[9].Status := '';
   OrderTable[9].CompleteTime := '';
   OrderTable[9].ErrorID := 0;
   OrderTable[10].OrderNo := 0;
   OrderTable[10].StepNo := 0;
   OrderTable[10].PlaceTime := '';
   OrderTable[10].Device := '';
   OrderTable[10].Sequence := 0;
   OrderTable[10].Status := '';
   OrderTable[10].CompleteTime := '';
   OrderTable[10].ErrorID := 0;
   OrderTable[11].OrderNo := 0;
   OrderTable[11].StepNo := 0;
   OrderTable[11].PlaceTime := '';
   OrderTable[11].Device := '';
   OrderTable[11].Sequence := 0;
   OrderTable[11].Status := '';
   OrderTable[11].CompleteTime := '';
   OrderTable[11].ErrorID := 0;
   OrderTable[12].OrderNo := 0;
   OrderTable[12].StepNo := 0;
   OrderTable[12].PlaceTime := '';
   OrderTable[12].Device := '';
   OrderTable[12].Sequence := 0;
   OrderTable[12].Status := '';
   OrderTable[12].CompleteTime := '';
   OrderTable[12].ErrorID := 0;
   OrderTable[13].OrderNo := 0;
   OrderTable[13].StepNo := 0;
   OrderTable[13].PlaceTime := '';
   OrderTable[13].Device := '';
   OrderTable[13].Sequence := 0;
   OrderTable[13].Status := '';
   OrderTable[13].CompleteTime := '';
   OrderTable[13].ErrorID := 0;
   OrderTable[14].OrderNo := 0;
   OrderTable[14].StepNo := 0;
   OrderTable[14].PlaceTime := '';
   OrderTable[14].Device := '';
   OrderTable[14].Sequence := 0;
   OrderTable[14].Status := '';
   OrderTable[14].CompleteTime := '';
   OrderTable[14].ErrorID := 0;
   OrderTable[15].OrderNo := 0;
   OrderTable[15].StepNo := 0;
   OrderTable[15].PlaceTime := '';
   OrderTable[15].Device := '';
   OrderTable[15].Sequence := 0;
   OrderTable[15].Status := '';
   OrderTable[15].CompleteTime := '';
   OrderTable[15].ErrorID := 0;
   OrderTable[16].OrderNo := 0;
   OrderTable[16].StepNo := 0;
   OrderTable[16].PlaceTime := '';
   OrderTable[16].Device := '';
   OrderTable[16].Sequence := 0;
   OrderTable[16].Status := '';
   OrderTable[16].CompleteTime := '';
   OrderTable[16].ErrorID := 0;
   OrderTable[17].OrderNo := 0;
   OrderTable[17].StepNo := 0;
   OrderTable[17].PlaceTime := '';
   OrderTable[17].Device := '';
   OrderTable[17].Sequence := 0;
   OrderTable[17].Status := '';
   OrderTable[17].CompleteTime := '';
   OrderTable[17].ErrorID := 0;
   OrderTable[18].OrderNo := 0;
   OrderTable[18].StepNo := 0;
   OrderTable[18].PlaceTime := '';
   OrderTable[18].Device := '';
   OrderTable[18].Sequence := 0;
   OrderTable[18].Status := '';
   OrderTable[18].CompleteTime := '';
   OrderTable[18].ErrorID := 0;
   OrderTable[19].OrderNo := 0;
   OrderTable[19].StepNo := 0;
   OrderTable[19].PlaceTime := '';
   OrderTable[19].Device := '';
   OrderTable[19].Sequence := 0;
   OrderTable[19].Status := '';
   OrderTable[19].CompleteTime := '';
   OrderTable[19].ErrorID := 0;
   OrderTable[20].OrderNo := 0;
   OrderTable[20].StepNo := 0;
   OrderTable[20].PlaceTime := '';
   OrderTable[20].Device := '';
   OrderTable[20].Sequence := 0;
   OrderTable[20].Status := '';
   OrderTable[20].CompleteTime := '';
   OrderTable[20].ErrorID := 0;
   OrderTable[21].OrderNo := 0;
   OrderTable[21].StepNo := 0;
   OrderTable[21].PlaceTime := '';
   OrderTable[21].Device := '';
   OrderTable[21].Sequence := 0;
   OrderTable[21].Status := '';
   OrderTable[21].CompleteTime := '';
   OrderTable[21].ErrorID := 0;
   OrderTable[22].OrderNo := 0;
   OrderTable[22].StepNo := 0;
   OrderTable[22].PlaceTime := '';
   OrderTable[22].Device := '';
   OrderTable[22].Sequence := 0;
   OrderTable[22].Status := '';
   OrderTable[22].CompleteTime := '';
   OrderTable[22].ErrorID := 0;
   OrderTable[23].OrderNo := 0;
   OrderTable[23].StepNo := 0;
   OrderTable[23].PlaceTime := '';
   OrderTable[23].Device := '';
   OrderTable[23].Sequence := 0;
   OrderTable[23].Status := '';
   OrderTable[23].CompleteTime := '';
   OrderTable[23].ErrorID := 0;
   OrderTable[24].OrderNo := 0;
   OrderTable[24].StepNo := 0;
   OrderTable[24].PlaceTime := '';
   OrderTable[24].Device := '';
   OrderTable[24].Sequence := 0;
   OrderTable[24].Status := '';
   OrderTable[24].CompleteTime := '';
   OrderTable[24].ErrorID := 0;
   OrderTable[25].OrderNo := 0;
   OrderTable[25].StepNo := 0;
   OrderTable[25].PlaceTime := '';
   OrderTable[25].Device := '';
   OrderTable[25].Sequence := 0;
   OrderTable[25].Status := '';
   OrderTable[25].CompleteTime := '';
   OrderTable[25].ErrorID := 0;
   OrderTable[26].OrderNo := 0;
   OrderTable[26].StepNo := 0;
   OrderTable[26].PlaceTime := '';
   OrderTable[26].Device := '';
   OrderTable[26].Sequence := 0;
   OrderTable[26].Status := '';
   OrderTable[26].CompleteTime := '';
   OrderTable[26].ErrorID := 0;
   OrderTable[27].OrderNo := 0;
   OrderTable[27].StepNo := 0;
   OrderTable[27].PlaceTime := '';
   OrderTable[27].Device := '';
   OrderTable[27].Sequence := 0;
   OrderTable[27].Status := '';
   OrderTable[27].CompleteTime := '';
   OrderTable[27].ErrorID := 0;
   OrderTable[28].OrderNo := 0;
   OrderTable[28].StepNo := 0;
   OrderTable[28].PlaceTime := '';
   OrderTable[28].Device := '';
   OrderTable[28].Sequence := 0;
   OrderTable[28].Status := '';
   OrderTable[28].CompleteTime := '';
   OrderTable[28].ErrorID := 0;
   OrderTable[29].OrderNo := 0;
   OrderTable[29].StepNo := 0;
   OrderTable[29].PlaceTime := '';
   OrderTable[29].Device := '';
   OrderTable[29].Sequence := 0;
   OrderTable[29].Status := '';
   OrderTable[29].CompleteTime := '';
   OrderTable[29].ErrorID := 0;
   OrderTable[30].OrderNo := 0;
   OrderTable[30].StepNo := 0;
   OrderTable[30].PlaceTime := '';
   OrderTable[30].Device := '';
   OrderTable[30].Sequence := 0;
   OrderTable[30].Status := '';
   OrderTable[30].CompleteTime := '';
   OrderTable[30].ErrorID := 0;
   OrderTable[31].OrderNo := 0;
   OrderTable[31].StepNo := 0;
   OrderTable[31].PlaceTime := '';
   OrderTable[31].Device := '';
   OrderTable[31].Sequence := 0;
   OrderTable[31].Status := '';
   OrderTable[31].CompleteTime := '';
   OrderTable[31].ErrorID := 0;
   OrderTable[32].OrderNo := 0;
   OrderTable[32].StepNo := 0;
   OrderTable[32].PlaceTime := '';
   OrderTable[32].Device := '';
   OrderTable[32].Sequence := 0;
   OrderTable[32].Status := '';
   OrderTable[32].CompleteTime := '';
   OrderTable[32].ErrorID := 0;
   OrderTable[33].OrderNo := 0;
   OrderTable[33].StepNo := 0;
   OrderTable[33].PlaceTime := '';
   OrderTable[33].Device := '';
   OrderTable[33].Sequence := 0;
   OrderTable[33].Status := '';
   OrderTable[33].CompleteTime := '';
   OrderTable[33].ErrorID := 0;
   OrderTable[34].OrderNo := 0;
   OrderTable[34].StepNo := 0;
   OrderTable[34].PlaceTime := '';
   OrderTable[34].Device := '';
   OrderTable[34].Sequence := 0;
   OrderTable[34].Status := '';
   OrderTable[34].CompleteTime := '';
   OrderTable[34].ErrorID := 0;
   OrderTable[35].OrderNo := 0;
   OrderTable[35].StepNo := 0;
   OrderTable[35].PlaceTime := '';
   OrderTable[35].Device := '';
   OrderTable[35].Sequence := 0;
   OrderTable[35].Status := '';
   OrderTable[35].CompleteTime := '';
   OrderTable[35].ErrorID := 0;
   OrderTable[36].OrderNo := 0;
   OrderTable[36].StepNo := 0;
   OrderTable[36].PlaceTime := '';
   OrderTable[36].Device := '';
   OrderTable[36].Sequence := 0;
   OrderTable[36].Status := '';
   OrderTable[36].CompleteTime := '';
   OrderTable[36].ErrorID := 0;
   OrderTable[37].OrderNo := 0;
   OrderTable[37].StepNo := 0;
   OrderTable[37].PlaceTime := '';
   OrderTable[37].Device := '';
   OrderTable[37].Sequence := 0;
   OrderTable[37].Status := '';
   OrderTable[37].CompleteTime := '';
   OrderTable[37].ErrorID := 0;
   OrderTable[38].OrderNo := 0;
   OrderTable[38].StepNo := 0;
   OrderTable[38].PlaceTime := '';
   OrderTable[38].Device := '';
   OrderTable[38].Sequence := 0;
   OrderTable[38].Status := '';
   OrderTable[38].CompleteTime := '';
   OrderTable[38].ErrorID := 0;
   OrderTable[39].OrderNo := 0;
   OrderTable[39].StepNo := 0;
   OrderTable[39].PlaceTime := '';
   OrderTable[39].Device := '';
   OrderTable[39].Sequence := 0;
   OrderTable[39].Status := '';
   OrderTable[39].CompleteTime := '';
   OrderTable[39].ErrorID := 0;
   OrderTable[40].OrderNo := 0;
   OrderTable[40].StepNo := 0;
   OrderTable[40].PlaceTime := '';
   OrderTable[40].Device := '';
   OrderTable[40].Sequence := 0;
   OrderTable[40].Status := '';
   OrderTable[40].CompleteTime := '';
   OrderTable[40].ErrorID := 0;
   OrderTable[41].OrderNo := 0;
   OrderTable[41].StepNo := 0;
   OrderTable[41].PlaceTime := '';
   OrderTable[41].Device := '';
   OrderTable[41].Sequence := 0;
   OrderTable[41].Status := '';
   OrderTable[41].CompleteTime := '';
   OrderTable[41].ErrorID := 0;
   OrderTable[42].OrderNo := 0;
   OrderTable[42].StepNo := 0;
   OrderTable[42].PlaceTime := '';
   OrderTable[42].Device := '';
   OrderTable[42].Sequence := 0;
   OrderTable[42].Status := '';
   OrderTable[42].CompleteTime := '';
   OrderTable[42].ErrorID := 0;
   OrderTable[43].OrderNo := 0;
   OrderTable[43].StepNo := 0;
   OrderTable[43].PlaceTime := '';
   OrderTable[43].Device := '';
   OrderTable[43].Sequence := 0;
   OrderTable[43].Status := '';
   OrderTable[43].CompleteTime := '';
   OrderTable[43].ErrorID := 0;
   OrderTable[44].OrderNo := 0;
   OrderTable[44].StepNo := 0;
   OrderTable[44].PlaceTime := '';
   OrderTable[44].Device := '';
   OrderTable[44].Sequence := 0;
   OrderTable[44].Status := '';
   OrderTable[44].CompleteTime := '';
   OrderTable[44].ErrorID := 0;
   OrderTable[45].OrderNo := 0;
   OrderTable[45].StepNo := 0;
   OrderTable[45].PlaceTime := '';
   OrderTable[45].Device := '';
   OrderTable[45].Sequence := 0;
   OrderTable[45].Status := '';
   OrderTable[45].CompleteTime := '';
   OrderTable[45].ErrorID := 0;
   OrderTable[46].OrderNo := 0;
   OrderTable[46].StepNo := 0;
   OrderTable[46].PlaceTime := '';
   OrderTable[46].Device := '';
   OrderTable[46].Sequence := 0;
   OrderTable[46].Status := '';
   OrderTable[46].CompleteTime := '';
   OrderTable[46].ErrorID := 0;
   OrderTable[47].OrderNo := 0;
   OrderTable[47].StepNo := 0;
   OrderTable[47].PlaceTime := '';
   OrderTable[47].Device := '';
   OrderTable[47].Sequence := 0;
   OrderTable[47].Status := '';
   OrderTable[47].CompleteTime := '';
   OrderTable[47].ErrorID := 0;
   OrderTable[48].OrderNo := 0;
   OrderTable[48].StepNo := 0;
   OrderTable[48].PlaceTime := '';
   OrderTable[48].Device := '';
   OrderTable[48].Sequence := 0;
   OrderTable[48].Status := '';
   OrderTable[48].CompleteTime := '';
   OrderTable[48].ErrorID := 0;
   OrderTable[49].OrderNo := 0;
   OrderTable[49].StepNo := 0;
   OrderTable[49].PlaceTime := '';
   OrderTable[49].Device := '';
   OrderTable[49].Sequence := 0;
   OrderTable[49].Status := '';
   OrderTable[49].CompleteTime := '';
   OrderTable[49].ErrorID := 0;
   OrderTable[50].OrderNo := 0;
   OrderTable[50].StepNo := 0;
   OrderTable[50].PlaceTime := '';
   OrderTable[50].Device := '';
   OrderTable[50].Sequence := 0;
   OrderTable[50].Status := '';
   OrderTable[50].CompleteTime := '';
   OrderTable[50].ErrorID := 0;
   OrderTable[51].OrderNo := 0;
   OrderTable[51].StepNo := 0;
   OrderTable[51].PlaceTime := '';
   OrderTable[51].Device := '';
   OrderTable[51].Sequence := 0;
   OrderTable[51].Status := '';
   OrderTable[51].CompleteTime := '';
   OrderTable[51].ErrorID := 0;
   OrderTable[52].OrderNo := 0;
   OrderTable[52].StepNo := 0;
   OrderTable[52].PlaceTime := '';
   OrderTable[52].Device := '';
   OrderTable[52].Sequence := 0;
   OrderTable[52].Status := '';
   OrderTable[52].CompleteTime := '';
   OrderTable[52].ErrorID := 0;
   OrderTable[53].OrderNo := 0;
   OrderTable[53].StepNo := 0;
   OrderTable[53].PlaceTime := '';
   OrderTable[53].Device := '';
   OrderTable[53].Sequence := 0;
   OrderTable[53].Status := '';
   OrderTable[53].CompleteTime := '';
   OrderTable[53].ErrorID := 0;
   OrderTable[54].OrderNo := 0;
   OrderTable[54].StepNo := 0;
   OrderTable[54].PlaceTime := '';
   OrderTable[54].Device := '';
   OrderTable[54].Sequence := 0;
   OrderTable[54].Status := '';
   OrderTable[54].CompleteTime := '';
   OrderTable[54].ErrorID := 0;
   OrderTable[55].OrderNo := 0;
   OrderTable[55].StepNo := 0;
   OrderTable[55].PlaceTime := '';
   OrderTable[55].Device := '';
   OrderTable[55].Sequence := 0;
   OrderTable[55].Status := '';
   OrderTable[55].CompleteTime := '';
   OrderTable[55].ErrorID := 0;
   OrderTable[56].OrderNo := 0;
   OrderTable[56].StepNo := 0;
   OrderTable[56].PlaceTime := '';
   OrderTable[56].Device := '';
   OrderTable[56].Sequence := 0;
   OrderTable[56].Status := '';
   OrderTable[56].CompleteTime := '';
   OrderTable[56].ErrorID := 0;
   OrderTable[57].OrderNo := 0;
   OrderTable[57].StepNo := 0;
   OrderTable[57].PlaceTime := '';
   OrderTable[57].Device := '';
   OrderTable[57].Sequence := 0;
   OrderTable[57].Status := '';
   OrderTable[57].CompleteTime := '';
   OrderTable[57].ErrorID := 0;
   OrderTable[58].OrderNo := 0;
   OrderTable[58].StepNo := 0;
   OrderTable[58].PlaceTime := '';
   OrderTable[58].Device := '';
   OrderTable[58].Sequence := 0;
   OrderTable[58].Status := '';
   OrderTable[58].CompleteTime := '';
   OrderTable[58].ErrorID := 0;
   OrderTable[59].OrderNo := 0;
   OrderTable[59].StepNo := 0;
   OrderTable[59].PlaceTime := '';
   OrderTable[59].Device := '';
   OrderTable[59].Sequence := 0;
   OrderTable[59].Status := '';
   OrderTable[59].CompleteTime := '';
   OrderTable[59].ErrorID := 0;
   OrderTable[60].OrderNo := 0;
   OrderTable[60].StepNo := 0;
   OrderTable[60].PlaceTime := '';
   OrderTable[60].Device := '';
   OrderTable[60].Sequence := 0;
   OrderTable[60].Status := '';
   OrderTable[60].CompleteTime := '';
   OrderTable[60].ErrorID := 0;
   OrderTable[61].OrderNo := 0;
   OrderTable[61].StepNo := 0;
   OrderTable[61].PlaceTime := '';
   OrderTable[61].Device := '';
   OrderTable[61].Sequence := 0;
   OrderTable[61].Status := '';
   OrderTable[61].CompleteTime := '';
   OrderTable[61].ErrorID := 0;
   OrderTable[62].OrderNo := 0;
   OrderTable[62].StepNo := 0;
   OrderTable[62].PlaceTime := '';
   OrderTable[62].Device := '';
   OrderTable[62].Sequence := 0;
   OrderTable[62].Status := '';
   OrderTable[62].CompleteTime := '';
   OrderTable[62].ErrorID := 0;
   OrderTable[63].OrderNo := 0;
   OrderTable[63].StepNo := 0;
   OrderTable[63].PlaceTime := '';
   OrderTable[63].Device := '';
   OrderTable[63].Sequence := 0;
   OrderTable[63].Status := '';
   OrderTable[63].CompleteTime := '';
   OrderTable[63].ErrorID := 0;
   OrderTable[64].OrderNo := 0;
   OrderTable[64].StepNo := 0;
   OrderTable[64].PlaceTime := '';
   OrderTable[64].Device := '';
   OrderTable[64].Sequence := 0;
   OrderTable[64].Status := '';
   OrderTable[64].CompleteTime := '';
   OrderTable[64].ErrorID := 0;
   OrderTable[65].OrderNo := 0;
   OrderTable[65].StepNo := 0;
   OrderTable[65].PlaceTime := '';
   OrderTable[65].Device := '';
   OrderTable[65].Sequence := 0;
   OrderTable[65].Status := '';
   OrderTable[65].CompleteTime := '';
   OrderTable[65].ErrorID := 0;
   OrderTable[66].OrderNo := 0;
   OrderTable[66].StepNo := 0;
   OrderTable[66].PlaceTime := '';
   OrderTable[66].Device := '';
   OrderTable[66].Sequence := 0;
   OrderTable[66].Status := '';
   OrderTable[66].CompleteTime := '';
   OrderTable[66].ErrorID := 0;
   OrderTable[67].OrderNo := 0;
   OrderTable[67].StepNo := 0;
   OrderTable[67].PlaceTime := '';
   OrderTable[67].Device := '';
   OrderTable[67].Sequence := 0;
   OrderTable[67].Status := '';
   OrderTable[67].CompleteTime := '';
   OrderTable[67].ErrorID := 0;
   OrderTable[68].OrderNo := 0;
   OrderTable[68].StepNo := 0;
   OrderTable[68].PlaceTime := '';
   OrderTable[68].Device := '';
   OrderTable[68].Sequence := 0;
   OrderTable[68].Status := '';
   OrderTable[68].CompleteTime := '';
   OrderTable[68].ErrorID := 0;
   OrderTable[69].OrderNo := 0;
   OrderTable[69].StepNo := 0;
   OrderTable[69].PlaceTime := '';
   OrderTable[69].Device := '';
   OrderTable[69].Sequence := 0;
   OrderTable[69].Status := '';
   OrderTable[69].CompleteTime := '';
   OrderTable[69].ErrorID := 0;
   OrderTable[70].OrderNo := 0;
   OrderTable[70].StepNo := 0;
   OrderTable[70].PlaceTime := '';
   OrderTable[70].Device := '';
   OrderTable[70].Sequence := 0;
   OrderTable[70].Status := '';
   OrderTable[70].CompleteTime := '';
   OrderTable[70].ErrorID := 0;
   OrderTable[71].OrderNo := 0;
   OrderTable[71].StepNo := 0;
   OrderTable[71].PlaceTime := '';
   OrderTable[71].Device := '';
   OrderTable[71].Sequence := 0;
   OrderTable[71].Status := '';
   OrderTable[71].CompleteTime := '';
   OrderTable[71].ErrorID := 0;
   OrderTable[72].OrderNo := 0;
   OrderTable[72].StepNo := 0;
   OrderTable[72].PlaceTime := '';
   OrderTable[72].Device := '';
   OrderTable[72].Sequence := 0;
   OrderTable[72].Status := '';
   OrderTable[72].CompleteTime := '';
   OrderTable[72].ErrorID := 0;
   OrderTable[73].OrderNo := 0;
   OrderTable[73].StepNo := 0;
   OrderTable[73].PlaceTime := '';
   OrderTable[73].Device := '';
   OrderTable[73].Sequence := 0;
   OrderTable[73].Status := '';
   OrderTable[73].CompleteTime := '';
   OrderTable[73].ErrorID := 0;
   OrderTable[74].OrderNo := 0;
   OrderTable[74].StepNo := 0;
   OrderTable[74].PlaceTime := '';
   OrderTable[74].Device := '';
   OrderTable[74].Sequence := 0;
   OrderTable[74].Status := '';
   OrderTable[74].CompleteTime := '';
   OrderTable[74].ErrorID := 0;
   OrderTable[75].OrderNo := 0;
   OrderTable[75].StepNo := 0;
   OrderTable[75].PlaceTime := '';
   OrderTable[75].Device := '';
   OrderTable[75].Sequence := 0;
   OrderTable[75].Status := '';
   OrderTable[75].CompleteTime := '';
   OrderTable[75].ErrorID := 0;
   OrderTable[76].OrderNo := 0;
   OrderTable[76].StepNo := 0;
   OrderTable[76].PlaceTime := '';
   OrderTable[76].Device := '';
   OrderTable[76].Sequence := 0;
   OrderTable[76].Status := '';
   OrderTable[76].CompleteTime := '';
   OrderTable[76].ErrorID := 0;
   OrderTable[77].OrderNo := 0;
   OrderTable[77].StepNo := 0;
   OrderTable[77].PlaceTime := '';
   OrderTable[77].Device := '';
   OrderTable[77].Sequence := 0;
   OrderTable[77].Status := '';
   OrderTable[77].CompleteTime := '';
   OrderTable[77].ErrorID := 0;
   OrderTable[78].OrderNo := 0;
   OrderTable[78].StepNo := 0;
   OrderTable[78].PlaceTime := '';
   OrderTable[78].Device := '';
   OrderTable[78].Sequence := 0;
   OrderTable[78].Status := '';
   OrderTable[78].CompleteTime := '';
   OrderTable[78].ErrorID := 0;
   OrderTable[79].OrderNo := 0;
   OrderTable[79].StepNo := 0;
   OrderTable[79].PlaceTime := '';
   OrderTable[79].Device := '';
   OrderTable[79].Sequence := 0;
   OrderTable[79].Status := '';
   OrderTable[79].CompleteTime := '';
   OrderTable[79].ErrorID := 0;
   OrderTable[80].OrderNo := 0;
   OrderTable[80].StepNo := 0;
   OrderTable[80].PlaceTime := '';
   OrderTable[80].Device := '';
   OrderTable[80].Sequence := 0;
   OrderTable[80].Status := '';
   OrderTable[80].CompleteTime := '';
   OrderTable[80].ErrorID := 0;
   OrderTable[81].OrderNo := 0;
   OrderTable[81].StepNo := 0;
   OrderTable[81].PlaceTime := '';
   OrderTable[81].Device := '';
   OrderTable[81].Sequence := 0;
   OrderTable[81].Status := '';
   OrderTable[81].CompleteTime := '';
   OrderTable[81].ErrorID := 0;
   OrderTable[82].OrderNo := 0;
   OrderTable[82].StepNo := 0;
   OrderTable[82].PlaceTime := '';
   OrderTable[82].Device := '';
   OrderTable[82].Sequence := 0;
   OrderTable[82].Status := '';
   OrderTable[82].CompleteTime := '';
   OrderTable[82].ErrorID := 0;
   OrderTable[83].OrderNo := 0;
   OrderTable[83].StepNo := 0;
   OrderTable[83].PlaceTime := '';
   OrderTable[83].Device := '';
   OrderTable[83].Sequence := 0;
   OrderTable[83].Status := '';
   OrderTable[83].CompleteTime := '';
   OrderTable[83].ErrorID := 0;
   OrderTable[84].OrderNo := 0;
   OrderTable[84].StepNo := 0;
   OrderTable[84].PlaceTime := '';
   OrderTable[84].Device := '';
   OrderTable[84].Sequence := 0;
   OrderTable[84].Status := '';
   OrderTable[84].CompleteTime := '';
   OrderTable[84].ErrorID := 0;
   OrderTable[85].OrderNo := 0;
   OrderTable[85].StepNo := 0;
   OrderTable[85].PlaceTime := '';
   OrderTable[85].Device := '';
   OrderTable[85].Sequence := 0;
   OrderTable[85].Status := '';
   OrderTable[85].CompleteTime := '';
   OrderTable[85].ErrorID := 0;
   OrderTable[86].OrderNo := 0;
   OrderTable[86].StepNo := 0;
   OrderTable[86].PlaceTime := '';
   OrderTable[86].Device := '';
   OrderTable[86].Sequence := 0;
   OrderTable[86].Status := '';
   OrderTable[86].CompleteTime := '';
   OrderTable[86].ErrorID := 0;
   OrderTable[87].OrderNo := 0;
   OrderTable[87].StepNo := 0;
   OrderTable[87].PlaceTime := '';
   OrderTable[87].Device := '';
   OrderTable[87].Sequence := 0;
   OrderTable[87].Status := '';
   OrderTable[87].CompleteTime := '';
   OrderTable[87].ErrorID := 0;
   OrderTable[88].OrderNo := 0;
   OrderTable[88].StepNo := 0;
   OrderTable[88].PlaceTime := '';
   OrderTable[88].Device := '';
   OrderTable[88].Sequence := 0;
   OrderTable[88].Status := '';
   OrderTable[88].CompleteTime := '';
   OrderTable[88].ErrorID := 0;
   OrderTable[89].OrderNo := 0;
   OrderTable[89].StepNo := 0;
   OrderTable[89].PlaceTime := '';
   OrderTable[89].Device := '';
   OrderTable[89].Sequence := 0;
   OrderTable[89].Status := '';
   OrderTable[89].CompleteTime := '';
   OrderTable[89].ErrorID := 0;
   OrderTable[90].OrderNo := 0;
   OrderTable[90].StepNo := 0;
   OrderTable[90].PlaceTime := '';
   OrderTable[90].Device := '';
   OrderTable[90].Sequence := 0;
   OrderTable[90].Status := '';
   OrderTable[90].CompleteTime := '';
   OrderTable[90].ErrorID := 0;
   OrderTable[91].OrderNo := 0;
   OrderTable[91].StepNo := 0;
   OrderTable[91].PlaceTime := '';
   OrderTable[91].Device := '';
   OrderTable[91].Sequence := 0;
   OrderTable[91].Status := '';
   OrderTable[91].CompleteTime := '';
   OrderTable[91].ErrorID := 0;
   OrderTable[92].OrderNo := 0;
   OrderTable[92].StepNo := 0;
   OrderTable[92].PlaceTime := '';
   OrderTable[92].Device := '';
   OrderTable[92].Sequence := 0;
   OrderTable[92].Status := '';
   OrderTable[92].CompleteTime := '';
   OrderTable[92].ErrorID := 0;
   OrderTable[93].OrderNo := 0;
   OrderTable[93].StepNo := 0;
   OrderTable[93].PlaceTime := '';
   OrderTable[93].Device := '';
   OrderTable[93].Sequence := 0;
   OrderTable[93].Status := '';
   OrderTable[93].CompleteTime := '';
   OrderTable[93].ErrorID := 0;
   OrderTable[94].OrderNo := 0;
   OrderTable[94].StepNo := 0;
   OrderTable[94].PlaceTime := '';
   OrderTable[94].Device := '';
   OrderTable[94].Sequence := 0;
   OrderTable[94].Status := '';
   OrderTable[94].CompleteTime := '';
   OrderTable[94].ErrorID := 0;
   OrderTable[95].OrderNo := 0;
   OrderTable[95].StepNo := 0;
   OrderTable[95].PlaceTime := '';
   OrderTable[95].Device := '';
   OrderTable[95].Sequence := 0;
   OrderTable[95].Status := '';
   OrderTable[95].CompleteTime := '';
   OrderTable[95].ErrorID := 0;
   OrderTable[96].OrderNo := 0;
   OrderTable[96].StepNo := 0;
   OrderTable[96].PlaceTime := '';
   OrderTable[96].Device := '';
   OrderTable[96].Sequence := 0;
   OrderTable[96].Status := '';
   OrderTable[96].CompleteTime := '';
   OrderTable[96].ErrorID := 0;
   OrderTable[97].OrderNo := 0;
   OrderTable[97].StepNo := 0;
   OrderTable[97].PlaceTime := '';
   OrderTable[97].Device := '';
   OrderTable[97].Sequence := 0;
   OrderTable[97].Status := '';
   OrderTable[97].CompleteTime := '';
   OrderTable[97].ErrorID := 0;
   OrderTable[98].OrderNo := 0;
   OrderTable[98].StepNo := 0;
   OrderTable[98].PlaceTime := '';
   OrderTable[98].Device := '';
   OrderTable[98].Sequence := 0;
   OrderTable[98].Status := '';
   OrderTable[98].CompleteTime := '';
   OrderTable[98].ErrorID := 0;
   OrderTable[99].OrderNo := 0;
   OrderTable[99].StepNo := 0;
   OrderTable[99].PlaceTime := '';
   OrderTable[99].Device := '';
   OrderTable[99].Sequence := 0;
   OrderTable[99].Status := '';
   OrderTable[99].CompleteTime := '';
   OrderTable[99].ErrorID := 0;
   StepTable[1].OrderNo := 0;
   StepTable[1].StepNo := 0;
   StepTable[1].PlaceTime := '';
   StepTable[1].Device := '';
   StepTable[1].Sequence := 0;
   StepTable[1].Status := '';
   StepTable[1].CompleteTime := '';
   StepTable[1].ErrorID := 0;
   StepTable[2].OrderNo := 0;
   StepTable[2].StepNo := 0;
   StepTable[2].PlaceTime := '';
   StepTable[2].Device := '';
   StepTable[2].Sequence := 0;
   StepTable[2].Status := '';
   StepTable[2].CompleteTime := '';
   StepTable[2].ErrorID := 0;
   StepTable[3].OrderNo := 0;
   StepTable[3].StepNo := 0;
   StepTable[3].PlaceTime := '';
   StepTable[3].Device := '';
   StepTable[3].Sequence := 0;
   StepTable[3].Status := '';
   StepTable[3].CompleteTime := '';
   StepTable[3].ErrorID := 0;
   StepTable[4].OrderNo := 0;
   StepTable[4].StepNo := 0;
   StepTable[4].PlaceTime := '';
   StepTable[4].Device := '';
   StepTable[4].Sequence := 0;
   StepTable[4].Status := '';
   StepTable[4].CompleteTime := '';
   StepTable[4].ErrorID := 0;
   StepTable[5].OrderNo := 0;
   StepTable[5].StepNo := 0;
   StepTable[5].PlaceTime := '';
   StepTable[5].Device := '';
   StepTable[5].Sequence := 0;
   StepTable[5].Status := '';
   StepTable[5].CompleteTime := '';
   StepTable[5].ErrorID := 0;
   StepTable[6].OrderNo := 0;
   StepTable[6].StepNo := 0;
   StepTable[6].PlaceTime := '';
   StepTable[6].Device := '';
   StepTable[6].Sequence := 0;
   StepTable[6].Status := '';
   StepTable[6].CompleteTime := '';
   StepTable[6].ErrorID := 0;
   StepTable[7].OrderNo := 0;
   StepTable[7].StepNo := 0;
   StepTable[7].PlaceTime := '';
   StepTable[7].Device := '';
   StepTable[7].Sequence := 0;
   StepTable[7].Status := '';
   StepTable[7].CompleteTime := '';
   StepTable[7].ErrorID := 0;
   StepTable[8].OrderNo := 0;
   StepTable[8].StepNo := 0;
   StepTable[8].PlaceTime := '';
   StepTable[8].Device := '';
   StepTable[8].Sequence := 0;
   StepTable[8].Status := '';
   StepTable[8].CompleteTime := '';
   StepTable[8].ErrorID := 0;
   StepTable[9].OrderNo := 0;
   StepTable[9].StepNo := 0;
   StepTable[9].PlaceTime := '';
   StepTable[9].Device := '';
   StepTable[9].Sequence := 0;
   StepTable[9].Status := '';
   StepTable[9].CompleteTime := '';
   StepTable[9].ErrorID := 0;
   StepTable[10].OrderNo := 0;
   StepTable[10].StepNo := 0;
   StepTable[10].PlaceTime := '';
   StepTable[10].Device := '';
   StepTable[10].Sequence := 0;
   StepTable[10].Status := '';
   StepTable[10].CompleteTime := '';
   StepTable[10].ErrorID := 0;
   StepTable[11].OrderNo := 0;
   StepTable[11].StepNo := 0;
   StepTable[11].PlaceTime := '';
   StepTable[11].Device := '';
   StepTable[11].Sequence := 0;
   StepTable[11].Status := '';
   StepTable[11].CompleteTime := '';
   StepTable[11].ErrorID := 0;
   StepTable[12].OrderNo := 0;
   StepTable[12].StepNo := 0;
   StepTable[12].PlaceTime := '';
   StepTable[12].Device := '';
   StepTable[12].Sequence := 0;
   StepTable[12].Status := '';
   StepTable[12].CompleteTime := '';
   StepTable[12].ErrorID := 0;
   StepTable[13].OrderNo := 0;
   StepTable[13].StepNo := 0;
   StepTable[13].PlaceTime := '';
   StepTable[13].Device := '';
   StepTable[13].Sequence := 0;
   StepTable[13].Status := '';
   StepTable[13].CompleteTime := '';
   StepTable[13].ErrorID := 0;
   StepTable[14].OrderNo := 0;
   StepTable[14].StepNo := 0;
   StepTable[14].PlaceTime := '';
   StepTable[14].Device := '';
   StepTable[14].Sequence := 0;
   StepTable[14].Status := '';
   StepTable[14].CompleteTime := '';
   StepTable[14].ErrorID := 0;
   StepTable[15].OrderNo := 0;
   StepTable[15].StepNo := 0;
   StepTable[15].PlaceTime := '';
   StepTable[15].Device := '';
   StepTable[15].Sequence := 0;
   StepTable[15].Status := '';
   StepTable[15].CompleteTime := '';
   StepTable[15].ErrorID := 0;
   StepTable[16].OrderNo := 0;
   StepTable[16].StepNo := 0;
   StepTable[16].PlaceTime := '';
   StepTable[16].Device := '';
   StepTable[16].Sequence := 0;
   StepTable[16].Status := '';
   StepTable[16].CompleteTime := '';
   StepTable[16].ErrorID := 0;
   StepTable[17].OrderNo := 0;
   StepTable[17].StepNo := 0;
   StepTable[17].PlaceTime := '';
   StepTable[17].Device := '';
   StepTable[17].Sequence := 0;
   StepTable[17].Status := '';
   StepTable[17].CompleteTime := '';
   StepTable[17].ErrorID := 0;
   StepTable[18].OrderNo := 0;
   StepTable[18].StepNo := 0;
   StepTable[18].PlaceTime := '';
   StepTable[18].Device := '';
   StepTable[18].Sequence := 0;
   StepTable[18].Status := '';
   StepTable[18].CompleteTime := '';
   StepTable[18].ErrorID := 0;
   StepTable[19].OrderNo := 0;
   StepTable[19].StepNo := 0;
   StepTable[19].PlaceTime := '';
   StepTable[19].Device := '';
   StepTable[19].Sequence := 0;
   StepTable[19].Status := '';
   StepTable[19].CompleteTime := '';
   StepTable[19].ErrorID := 0;
   StepTable[20].OrderNo := 0;
   StepTable[20].StepNo := 0;
   StepTable[20].PlaceTime := '';
   StepTable[20].Device := '';
   StepTable[20].Sequence := 0;
   StepTable[20].Status := '';
   StepTable[20].CompleteTime := '';
   StepTable[20].ErrorID := 0;
   CarParked_Confirm := FALSE;
   Running := FALSE;
   IDLE := TRUE;
   Error := FALSE;
   State := 0;
   ResetError := FALSE;
   Ready := TRUE;
   Selected := TRUE;
   Auto_Man := TRUE;
   Paused := FALSE;

END_DATA_BLOCK

DATA_BLOCK "Auto_Test_1_DB"
{ S7_Optimized_Access := 'TRUE' }
VERSION : 0.1
NON_RETAIN
"Auto_Test"

BEGIN

END_DATA_BLOCK

DATA_BLOCK "Auto_Test_3_DB"
{ S7_Optimized_Access := 'TRUE' }
VERSION : 0.1
NON_RETAIN
"Auto_Test"

BEGIN

END_DATA_BLOCK

DATA_BLOCK "System_DB_1"
{ S7_Optimized_Access := 'TRUE' }
VERSION : 0.1
NON_RETAIN
"System_UDT"

BEGIN
   Id := 1;
   CancelOrders := FALSE;
   PauseOrders := FALSE;
   ResumeOrders := FALSE;
   OrderSent := FALSE;
   CurrentOrder := 0;
   NextOrder := 1;
   OrderTable[0].OrderNo := 0;
   OrderTable[0].StepNo := 256;
   OrderTable[0].PlaceTime := '';
   OrderTable[0].Device := '';
   OrderTable[0].Sequence := 0;
   OrderTable[0].Status := 'Error';
   OrderTable[0].CompleteTime := '06/10/2022 08:58:15';
   OrderTable[0].ErrorID := 0;
   OrderTable[1].OrderNo := 0;
   OrderTable[1].StepNo := 0;
   OrderTable[1].PlaceTime := '';
   OrderTable[1].Device := '';
   OrderTable[1].Sequence := 0;
   OrderTable[1].Status := '';
   OrderTable[1].CompleteTime := '';
   OrderTable[1].ErrorID := 0;
   OrderTable[2].OrderNo := 0;
   OrderTable[2].StepNo := 0;
   OrderTable[2].PlaceTime := '';
   OrderTable[2].Device := '';
   OrderTable[2].Sequence := 0;
   OrderTable[2].Status := '';
   OrderTable[2].CompleteTime := '';
   OrderTable[2].ErrorID := 0;
   OrderTable[3].OrderNo := 0;
   OrderTable[3].StepNo := 0;
   OrderTable[3].PlaceTime := '';
   OrderTable[3].Device := '';
   OrderTable[3].Sequence := 0;
   OrderTable[3].Status := '';
   OrderTable[3].CompleteTime := '';
   OrderTable[3].ErrorID := 0;
   OrderTable[4].OrderNo := 0;
   OrderTable[4].StepNo := 0;
   OrderTable[4].PlaceTime := '';
   OrderTable[4].Device := '';
   OrderTable[4].Sequence := 0;
   OrderTable[4].Status := '';
   OrderTable[4].CompleteTime := '';
   OrderTable[4].ErrorID := 0;
   OrderTable[5].OrderNo := 0;
   OrderTable[5].StepNo := 0;
   OrderTable[5].PlaceTime := '';
   OrderTable[5].Device := '';
   OrderTable[5].Sequence := 0;
   OrderTable[5].Status := '';
   OrderTable[5].CompleteTime := '';
   OrderTable[5].ErrorID := 0;
   OrderTable[6].OrderNo := 0;
   OrderTable[6].StepNo := 0;
   OrderTable[6].PlaceTime := '';
   OrderTable[6].Device := '';
   OrderTable[6].Sequence := 0;
   OrderTable[6].Status := '';
   OrderTable[6].CompleteTime := '';
   OrderTable[6].ErrorID := 0;
   OrderTable[7].OrderNo := 0;
   OrderTable[7].StepNo := 0;
   OrderTable[7].PlaceTime := '';
   OrderTable[7].Device := '';
   OrderTable[7].Sequence := 0;
   OrderTable[7].Status := '';
   OrderTable[7].CompleteTime := '';
   OrderTable[7].ErrorID := 0;
   OrderTable[8].OrderNo := 0;
   OrderTable[8].StepNo := 0;
   OrderTable[8].PlaceTime := '';
   OrderTable[8].Device := '';
   OrderTable[8].Sequence := 0;
   OrderTable[8].Status := '';
   OrderTable[8].CompleteTime := '';
   OrderTable[8].ErrorID := 0;
   OrderTable[9].OrderNo := 0;
   OrderTable[9].StepNo := 0;
   OrderTable[9].PlaceTime := '';
   OrderTable[9].Device := '';
   OrderTable[9].Sequence := 0;
   OrderTable[9].Status := '';
   OrderTable[9].CompleteTime := '';
   OrderTable[9].ErrorID := 0;
   OrderTable[10].OrderNo := 0;
   OrderTable[10].StepNo := 0;
   OrderTable[10].PlaceTime := '';
   OrderTable[10].Device := '';
   OrderTable[10].Sequence := 0;
   OrderTable[10].Status := '';
   OrderTable[10].CompleteTime := '';
   OrderTable[10].ErrorID := 0;
   OrderTable[11].OrderNo := 0;
   OrderTable[11].StepNo := 0;
   OrderTable[11].PlaceTime := '';
   OrderTable[11].Device := '';
   OrderTable[11].Sequence := 0;
   OrderTable[11].Status := '';
   OrderTable[11].CompleteTime := '';
   OrderTable[11].ErrorID := 0;
   OrderTable[12].OrderNo := 0;
   OrderTable[12].StepNo := 0;
   OrderTable[12].PlaceTime := '';
   OrderTable[12].Device := '';
   OrderTable[12].Sequence := 0;
   OrderTable[12].Status := '';
   OrderTable[12].CompleteTime := '';
   OrderTable[12].ErrorID := 0;
   OrderTable[13].OrderNo := 0;
   OrderTable[13].StepNo := 0;
   OrderTable[13].PlaceTime := '';
   OrderTable[13].Device := '';
   OrderTable[13].Sequence := 0;
   OrderTable[13].Status := '';
   OrderTable[13].CompleteTime := '';
   OrderTable[13].ErrorID := 0;
   OrderTable[14].OrderNo := 0;
   OrderTable[14].StepNo := 0;
   OrderTable[14].PlaceTime := '';
   OrderTable[14].Device := '';
   OrderTable[14].Sequence := 0;
   OrderTable[14].Status := '';
   OrderTable[14].CompleteTime := '';
   OrderTable[14].ErrorID := 0;
   OrderTable[15].OrderNo := 0;
   OrderTable[15].StepNo := 0;
   OrderTable[15].PlaceTime := '';
   OrderTable[15].Device := '';
   OrderTable[15].Sequence := 0;
   OrderTable[15].Status := '';
   OrderTable[15].CompleteTime := '';
   OrderTable[15].ErrorID := 0;
   OrderTable[16].OrderNo := 0;
   OrderTable[16].StepNo := 0;
   OrderTable[16].PlaceTime := '';
   OrderTable[16].Device := '';
   OrderTable[16].Sequence := 0;
   OrderTable[16].Status := '';
   OrderTable[16].CompleteTime := '';
   OrderTable[16].ErrorID := 0;
   OrderTable[17].OrderNo := 0;
   OrderTable[17].StepNo := 0;
   OrderTable[17].PlaceTime := '';
   OrderTable[17].Device := '';
   OrderTable[17].Sequence := 0;
   OrderTable[17].Status := '';
   OrderTable[17].CompleteTime := '';
   OrderTable[17].ErrorID := 0;
   OrderTable[18].OrderNo := 0;
   OrderTable[18].StepNo := 0;
   OrderTable[18].PlaceTime := '';
   OrderTable[18].Device := '';
   OrderTable[18].Sequence := 0;
   OrderTable[18].Status := '';
   OrderTable[18].CompleteTime := '';
   OrderTable[18].ErrorID := 0;
   OrderTable[19].OrderNo := 0;
   OrderTable[19].StepNo := 0;
   OrderTable[19].PlaceTime := '';
   OrderTable[19].Device := '';
   OrderTable[19].Sequence := 0;
   OrderTable[19].Status := '';
   OrderTable[19].CompleteTime := '';
   OrderTable[19].ErrorID := 0;
   OrderTable[20].OrderNo := 0;
   OrderTable[20].StepNo := 0;
   OrderTable[20].PlaceTime := '';
   OrderTable[20].Device := '';
   OrderTable[20].Sequence := 0;
   OrderTable[20].Status := '';
   OrderTable[20].CompleteTime := '';
   OrderTable[20].ErrorID := 0;
   OrderTable[21].OrderNo := 0;
   OrderTable[21].StepNo := 0;
   OrderTable[21].PlaceTime := '';
   OrderTable[21].Device := '';
   OrderTable[21].Sequence := 0;
   OrderTable[21].Status := '';
   OrderTable[21].CompleteTime := '';
   OrderTable[21].ErrorID := 0;
   OrderTable[22].OrderNo := 0;
   OrderTable[22].StepNo := 0;
   OrderTable[22].PlaceTime := '';
   OrderTable[22].Device := '';
   OrderTable[22].Sequence := 0;
   OrderTable[22].Status := '';
   OrderTable[22].CompleteTime := '';
   OrderTable[22].ErrorID := 0;
   OrderTable[23].OrderNo := 0;
   OrderTable[23].StepNo := 0;
   OrderTable[23].PlaceTime := '';
   OrderTable[23].Device := '';
   OrderTable[23].Sequence := 0;
   OrderTable[23].Status := '';
   OrderTable[23].CompleteTime := '';
   OrderTable[23].ErrorID := 0;
   OrderTable[24].OrderNo := 0;
   OrderTable[24].StepNo := 0;
   OrderTable[24].PlaceTime := '';
   OrderTable[24].Device := '';
   OrderTable[24].Sequence := 0;
   OrderTable[24].Status := '';
   OrderTable[24].CompleteTime := '';
   OrderTable[24].ErrorID := 0;
   OrderTable[25].OrderNo := 0;
   OrderTable[25].StepNo := 0;
   OrderTable[25].PlaceTime := '';
   OrderTable[25].Device := '';
   OrderTable[25].Sequence := 0;
   OrderTable[25].Status := '';
   OrderTable[25].CompleteTime := '';
   OrderTable[25].ErrorID := 0;
   OrderTable[26].OrderNo := 0;
   OrderTable[26].StepNo := 0;
   OrderTable[26].PlaceTime := '';
   OrderTable[26].Device := '';
   OrderTable[26].Sequence := 0;
   OrderTable[26].Status := '';
   OrderTable[26].CompleteTime := '';
   OrderTable[26].ErrorID := 0;
   OrderTable[27].OrderNo := 0;
   OrderTable[27].StepNo := 0;
   OrderTable[27].PlaceTime := '';
   OrderTable[27].Device := '';
   OrderTable[27].Sequence := 0;
   OrderTable[27].Status := '';
   OrderTable[27].CompleteTime := '';
   OrderTable[27].ErrorID := 0;
   OrderTable[28].OrderNo := 0;
   OrderTable[28].StepNo := 0;
   OrderTable[28].PlaceTime := '';
   OrderTable[28].Device := '';
   OrderTable[28].Sequence := 0;
   OrderTable[28].Status := '';
   OrderTable[28].CompleteTime := '';
   OrderTable[28].ErrorID := 0;
   OrderTable[29].OrderNo := 0;
   OrderTable[29].StepNo := 0;
   OrderTable[29].PlaceTime := '';
   OrderTable[29].Device := '';
   OrderTable[29].Sequence := 0;
   OrderTable[29].Status := '';
   OrderTable[29].CompleteTime := '';
   OrderTable[29].ErrorID := 0;
   OrderTable[30].OrderNo := 0;
   OrderTable[30].StepNo := 0;
   OrderTable[30].PlaceTime := '';
   OrderTable[30].Device := '';
   OrderTable[30].Sequence := 0;
   OrderTable[30].Status := '';
   OrderTable[30].CompleteTime := '';
   OrderTable[30].ErrorID := 0;
   OrderTable[31].OrderNo := 0;
   OrderTable[31].StepNo := 0;
   OrderTable[31].PlaceTime := '';
   OrderTable[31].Device := '';
   OrderTable[31].Sequence := 0;
   OrderTable[31].Status := '';
   OrderTable[31].CompleteTime := '';
   OrderTable[31].ErrorID := 0;
   OrderTable[32].OrderNo := 0;
   OrderTable[32].StepNo := 0;
   OrderTable[32].PlaceTime := '';
   OrderTable[32].Device := '';
   OrderTable[32].Sequence := 0;
   OrderTable[32].Status := '';
   OrderTable[32].CompleteTime := '';
   OrderTable[32].ErrorID := 0;
   OrderTable[33].OrderNo := 0;
   OrderTable[33].StepNo := 0;
   OrderTable[33].PlaceTime := '';
   OrderTable[33].Device := '';
   OrderTable[33].Sequence := 0;
   OrderTable[33].Status := '';
   OrderTable[33].CompleteTime := '';
   OrderTable[33].ErrorID := 0;
   OrderTable[34].OrderNo := 0;
   OrderTable[34].StepNo := 0;
   OrderTable[34].PlaceTime := '';
   OrderTable[34].Device := '';
   OrderTable[34].Sequence := 0;
   OrderTable[34].Status := '';
   OrderTable[34].CompleteTime := '';
   OrderTable[34].ErrorID := 0;
   OrderTable[35].OrderNo := 0;
   OrderTable[35].StepNo := 0;
   OrderTable[35].PlaceTime := '';
   OrderTable[35].Device := '';
   OrderTable[35].Sequence := 0;
   OrderTable[35].Status := '';
   OrderTable[35].CompleteTime := '';
   OrderTable[35].ErrorID := 0;
   OrderTable[36].OrderNo := 0;
   OrderTable[36].StepNo := 0;
   OrderTable[36].PlaceTime := '';
   OrderTable[36].Device := '';
   OrderTable[36].Sequence := 0;
   OrderTable[36].Status := '';
   OrderTable[36].CompleteTime := '';
   OrderTable[36].ErrorID := 0;
   OrderTable[37].OrderNo := 0;
   OrderTable[37].StepNo := 0;
   OrderTable[37].PlaceTime := '';
   OrderTable[37].Device := '';
   OrderTable[37].Sequence := 0;
   OrderTable[37].Status := '';
   OrderTable[37].CompleteTime := '';
   OrderTable[37].ErrorID := 0;
   OrderTable[38].OrderNo := 0;
   OrderTable[38].StepNo := 0;
   OrderTable[38].PlaceTime := '';
   OrderTable[38].Device := '';
   OrderTable[38].Sequence := 0;
   OrderTable[38].Status := '';
   OrderTable[38].CompleteTime := '';
   OrderTable[38].ErrorID := 0;
   OrderTable[39].OrderNo := 0;
   OrderTable[39].StepNo := 0;
   OrderTable[39].PlaceTime := '';
   OrderTable[39].Device := '';
   OrderTable[39].Sequence := 0;
   OrderTable[39].Status := '';
   OrderTable[39].CompleteTime := '';
   OrderTable[39].ErrorID := 0;
   OrderTable[40].OrderNo := 0;
   OrderTable[40].StepNo := 0;
   OrderTable[40].PlaceTime := '';
   OrderTable[40].Device := '';
   OrderTable[40].Sequence := 0;
   OrderTable[40].Status := '';
   OrderTable[40].CompleteTime := '';
   OrderTable[40].ErrorID := 0;
   OrderTable[41].OrderNo := 0;
   OrderTable[41].StepNo := 0;
   OrderTable[41].PlaceTime := '';
   OrderTable[41].Device := '';
   OrderTable[41].Sequence := 0;
   OrderTable[41].Status := '';
   OrderTable[41].CompleteTime := '';
   OrderTable[41].ErrorID := 0;
   OrderTable[42].OrderNo := 0;
   OrderTable[42].StepNo := 0;
   OrderTable[42].PlaceTime := '';
   OrderTable[42].Device := '';
   OrderTable[42].Sequence := 0;
   OrderTable[42].Status := '';
   OrderTable[42].CompleteTime := '';
   OrderTable[42].ErrorID := 0;
   OrderTable[43].OrderNo := 0;
   OrderTable[43].StepNo := 0;
   OrderTable[43].PlaceTime := '';
   OrderTable[43].Device := '';
   OrderTable[43].Sequence := 0;
   OrderTable[43].Status := '';
   OrderTable[43].CompleteTime := '';
   OrderTable[43].ErrorID := 0;
   OrderTable[44].OrderNo := 0;
   OrderTable[44].StepNo := 0;
   OrderTable[44].PlaceTime := '';
   OrderTable[44].Device := '';
   OrderTable[44].Sequence := 0;
   OrderTable[44].Status := '';
   OrderTable[44].CompleteTime := '';
   OrderTable[44].ErrorID := 0;
   OrderTable[45].OrderNo := 0;
   OrderTable[45].StepNo := 0;
   OrderTable[45].PlaceTime := '';
   OrderTable[45].Device := '';
   OrderTable[45].Sequence := 0;
   OrderTable[45].Status := '';
   OrderTable[45].CompleteTime := '';
   OrderTable[45].ErrorID := 0;
   OrderTable[46].OrderNo := 0;
   OrderTable[46].StepNo := 0;
   OrderTable[46].PlaceTime := '';
   OrderTable[46].Device := '';
   OrderTable[46].Sequence := 0;
   OrderTable[46].Status := '';
   OrderTable[46].CompleteTime := '';
   OrderTable[46].ErrorID := 0;
   OrderTable[47].OrderNo := 0;
   OrderTable[47].StepNo := 0;
   OrderTable[47].PlaceTime := '';
   OrderTable[47].Device := '';
   OrderTable[47].Sequence := 0;
   OrderTable[47].Status := '';
   OrderTable[47].CompleteTime := '';
   OrderTable[47].ErrorID := 0;
   OrderTable[48].OrderNo := 0;
   OrderTable[48].StepNo := 0;
   OrderTable[48].PlaceTime := '';
   OrderTable[48].Device := '';
   OrderTable[48].Sequence := 0;
   OrderTable[48].Status := '';
   OrderTable[48].CompleteTime := '';
   OrderTable[48].ErrorID := 0;
   OrderTable[49].OrderNo := 0;
   OrderTable[49].StepNo := 0;
   OrderTable[49].PlaceTime := '';
   OrderTable[49].Device := '';
   OrderTable[49].Sequence := 0;
   OrderTable[49].Status := '';
   OrderTable[49].CompleteTime := '';
   OrderTable[49].ErrorID := 0;
   OrderTable[50].OrderNo := 0;
   OrderTable[50].StepNo := 0;
   OrderTable[50].PlaceTime := '';
   OrderTable[50].Device := '';
   OrderTable[50].Sequence := 0;
   OrderTable[50].Status := '';
   OrderTable[50].CompleteTime := '';
   OrderTable[50].ErrorID := 0;
   OrderTable[51].OrderNo := 0;
   OrderTable[51].StepNo := 0;
   OrderTable[51].PlaceTime := '';
   OrderTable[51].Device := '';
   OrderTable[51].Sequence := 0;
   OrderTable[51].Status := '';
   OrderTable[51].CompleteTime := '';
   OrderTable[51].ErrorID := 0;
   OrderTable[52].OrderNo := 0;
   OrderTable[52].StepNo := 0;
   OrderTable[52].PlaceTime := '';
   OrderTable[52].Device := '';
   OrderTable[52].Sequence := 0;
   OrderTable[52].Status := '';
   OrderTable[52].CompleteTime := '';
   OrderTable[52].ErrorID := 0;
   OrderTable[53].OrderNo := 0;
   OrderTable[53].StepNo := 0;
   OrderTable[53].PlaceTime := '';
   OrderTable[53].Device := '';
   OrderTable[53].Sequence := 0;
   OrderTable[53].Status := '';
   OrderTable[53].CompleteTime := '';
   OrderTable[53].ErrorID := 0;
   OrderTable[54].OrderNo := 0;
   OrderTable[54].StepNo := 0;
   OrderTable[54].PlaceTime := '';
   OrderTable[54].Device := '';
   OrderTable[54].Sequence := 0;
   OrderTable[54].Status := '';
   OrderTable[54].CompleteTime := '';
   OrderTable[54].ErrorID := 0;
   OrderTable[55].OrderNo := 0;
   OrderTable[55].StepNo := 0;
   OrderTable[55].PlaceTime := '';
   OrderTable[55].Device := '';
   OrderTable[55].Sequence := 0;
   OrderTable[55].Status := '';
   OrderTable[55].CompleteTime := '';
   OrderTable[55].ErrorID := 0;
   OrderTable[56].OrderNo := 0;
   OrderTable[56].StepNo := 0;
   OrderTable[56].PlaceTime := '';
   OrderTable[56].Device := '';
   OrderTable[56].Sequence := 0;
   OrderTable[56].Status := '';
   OrderTable[56].CompleteTime := '';
   OrderTable[56].ErrorID := 0;
   OrderTable[57].OrderNo := 0;
   OrderTable[57].StepNo := 0;
   OrderTable[57].PlaceTime := '';
   OrderTable[57].Device := '';
   OrderTable[57].Sequence := 0;
   OrderTable[57].Status := '';
   OrderTable[57].CompleteTime := '';
   OrderTable[57].ErrorID := 0;
   OrderTable[58].OrderNo := 0;
   OrderTable[58].StepNo := 0;
   OrderTable[58].PlaceTime := '';
   OrderTable[58].Device := '';
   OrderTable[58].Sequence := 0;
   OrderTable[58].Status := '';
   OrderTable[58].CompleteTime := '';
   OrderTable[58].ErrorID := 0;
   OrderTable[59].OrderNo := 0;
   OrderTable[59].StepNo := 0;
   OrderTable[59].PlaceTime := '';
   OrderTable[59].Device := '';
   OrderTable[59].Sequence := 0;
   OrderTable[59].Status := '';
   OrderTable[59].CompleteTime := '';
   OrderTable[59].ErrorID := 0;
   OrderTable[60].OrderNo := 0;
   OrderTable[60].StepNo := 0;
   OrderTable[60].PlaceTime := '';
   OrderTable[60].Device := '';
   OrderTable[60].Sequence := 0;
   OrderTable[60].Status := '';
   OrderTable[60].CompleteTime := '';
   OrderTable[60].ErrorID := 0;
   OrderTable[61].OrderNo := 0;
   OrderTable[61].StepNo := 0;
   OrderTable[61].PlaceTime := '';
   OrderTable[61].Device := '';
   OrderTable[61].Sequence := 0;
   OrderTable[61].Status := '';
   OrderTable[61].CompleteTime := '';
   OrderTable[61].ErrorID := 0;
   OrderTable[62].OrderNo := 0;
   OrderTable[62].StepNo := 0;
   OrderTable[62].PlaceTime := '';
   OrderTable[62].Device := '';
   OrderTable[62].Sequence := 0;
   OrderTable[62].Status := '';
   OrderTable[62].CompleteTime := '';
   OrderTable[62].ErrorID := 0;
   OrderTable[63].OrderNo := 0;
   OrderTable[63].StepNo := 0;
   OrderTable[63].PlaceTime := '';
   OrderTable[63].Device := '';
   OrderTable[63].Sequence := 0;
   OrderTable[63].Status := '';
   OrderTable[63].CompleteTime := '';
   OrderTable[63].ErrorID := 0;
   OrderTable[64].OrderNo := 0;
   OrderTable[64].StepNo := 0;
   OrderTable[64].PlaceTime := '';
   OrderTable[64].Device := '';
   OrderTable[64].Sequence := 0;
   OrderTable[64].Status := '';
   OrderTable[64].CompleteTime := '';
   OrderTable[64].ErrorID := 0;
   OrderTable[65].OrderNo := 0;
   OrderTable[65].StepNo := 0;
   OrderTable[65].PlaceTime := '';
   OrderTable[65].Device := '';
   OrderTable[65].Sequence := 0;
   OrderTable[65].Status := '';
   OrderTable[65].CompleteTime := '';
   OrderTable[65].ErrorID := 0;
   OrderTable[66].OrderNo := 0;
   OrderTable[66].StepNo := 0;
   OrderTable[66].PlaceTime := '';
   OrderTable[66].Device := '';
   OrderTable[66].Sequence := 0;
   OrderTable[66].Status := '';
   OrderTable[66].CompleteTime := '';
   OrderTable[66].ErrorID := 0;
   OrderTable[67].OrderNo := 0;
   OrderTable[67].StepNo := 0;
   OrderTable[67].PlaceTime := '';
   OrderTable[67].Device := '';
   OrderTable[67].Sequence := 0;
   OrderTable[67].Status := '';
   OrderTable[67].CompleteTime := '';
   OrderTable[67].ErrorID := 0;
   OrderTable[68].OrderNo := 0;
   OrderTable[68].StepNo := 0;
   OrderTable[68].PlaceTime := '';
   OrderTable[68].Device := '';
   OrderTable[68].Sequence := 0;
   OrderTable[68].Status := '';
   OrderTable[68].CompleteTime := '';
   OrderTable[68].ErrorID := 0;
   OrderTable[69].OrderNo := 0;
   OrderTable[69].StepNo := 0;
   OrderTable[69].PlaceTime := '';
   OrderTable[69].Device := '';
   OrderTable[69].Sequence := 0;
   OrderTable[69].Status := '';
   OrderTable[69].CompleteTime := '';
   OrderTable[69].ErrorID := 0;
   OrderTable[70].OrderNo := 0;
   OrderTable[70].StepNo := 0;
   OrderTable[70].PlaceTime := '';
   OrderTable[70].Device := '';
   OrderTable[70].Sequence := 0;
   OrderTable[70].Status := '';
   OrderTable[70].CompleteTime := '';
   OrderTable[70].ErrorID := 0;
   OrderTable[71].OrderNo := 0;
   OrderTable[71].StepNo := 0;
   OrderTable[71].PlaceTime := '';
   OrderTable[71].Device := '';
   OrderTable[71].Sequence := 0;
   OrderTable[71].Status := '';
   OrderTable[71].CompleteTime := '';
   OrderTable[71].ErrorID := 0;
   OrderTable[72].OrderNo := 0;
   OrderTable[72].StepNo := 0;
   OrderTable[72].PlaceTime := '';
   OrderTable[72].Device := '';
   OrderTable[72].Sequence := 0;
   OrderTable[72].Status := '';
   OrderTable[72].CompleteTime := '';
   OrderTable[72].ErrorID := 0;
   OrderTable[73].OrderNo := 0;
   OrderTable[73].StepNo := 0;
   OrderTable[73].PlaceTime := '';
   OrderTable[73].Device := '';
   OrderTable[73].Sequence := 0;
   OrderTable[73].Status := '';
   OrderTable[73].CompleteTime := '';
   OrderTable[73].ErrorID := 0;
   OrderTable[74].OrderNo := 0;
   OrderTable[74].StepNo := 0;
   OrderTable[74].PlaceTime := '';
   OrderTable[74].Device := '';
   OrderTable[74].Sequence := 0;
   OrderTable[74].Status := '';
   OrderTable[74].CompleteTime := '';
   OrderTable[74].ErrorID := 0;
   OrderTable[75].OrderNo := 0;
   OrderTable[75].StepNo := 0;
   OrderTable[75].PlaceTime := '';
   OrderTable[75].Device := '';
   OrderTable[75].Sequence := 0;
   OrderTable[75].Status := '';
   OrderTable[75].CompleteTime := '';
   OrderTable[75].ErrorID := 0;
   OrderTable[76].OrderNo := 0;
   OrderTable[76].StepNo := 0;
   OrderTable[76].PlaceTime := '';
   OrderTable[76].Device := '';
   OrderTable[76].Sequence := 0;
   OrderTable[76].Status := '';
   OrderTable[76].CompleteTime := '';
   OrderTable[76].ErrorID := 0;
   OrderTable[77].OrderNo := 0;
   OrderTable[77].StepNo := 0;
   OrderTable[77].PlaceTime := '';
   OrderTable[77].Device := '';
   OrderTable[77].Sequence := 0;
   OrderTable[77].Status := '';
   OrderTable[77].CompleteTime := '';
   OrderTable[77].ErrorID := 0;
   OrderTable[78].OrderNo := 0;
   OrderTable[78].StepNo := 0;
   OrderTable[78].PlaceTime := '';
   OrderTable[78].Device := '';
   OrderTable[78].Sequence := 0;
   OrderTable[78].Status := '';
   OrderTable[78].CompleteTime := '';
   OrderTable[78].ErrorID := 0;
   OrderTable[79].OrderNo := 0;
   OrderTable[79].StepNo := 0;
   OrderTable[79].PlaceTime := '';
   OrderTable[79].Device := '';
   OrderTable[79].Sequence := 0;
   OrderTable[79].Status := '';
   OrderTable[79].CompleteTime := '';
   OrderTable[79].ErrorID := 0;
   OrderTable[80].OrderNo := 0;
   OrderTable[80].StepNo := 0;
   OrderTable[80].PlaceTime := '';
   OrderTable[80].Device := '';
   OrderTable[80].Sequence := 0;
   OrderTable[80].Status := '';
   OrderTable[80].CompleteTime := '';
   OrderTable[80].ErrorID := 0;
   OrderTable[81].OrderNo := 0;
   OrderTable[81].StepNo := 0;
   OrderTable[81].PlaceTime := '';
   OrderTable[81].Device := '';
   OrderTable[81].Sequence := 0;
   OrderTable[81].Status := '';
   OrderTable[81].CompleteTime := '';
   OrderTable[81].ErrorID := 0;
   OrderTable[82].OrderNo := 0;
   OrderTable[82].StepNo := 0;
   OrderTable[82].PlaceTime := '';
   OrderTable[82].Device := '';
   OrderTable[82].Sequence := 0;
   OrderTable[82].Status := '';
   OrderTable[82].CompleteTime := '';
   OrderTable[82].ErrorID := 0;
   OrderTable[83].OrderNo := 0;
   OrderTable[83].StepNo := 0;
   OrderTable[83].PlaceTime := '';
   OrderTable[83].Device := '';
   OrderTable[83].Sequence := 0;
   OrderTable[83].Status := '';
   OrderTable[83].CompleteTime := '';
   OrderTable[83].ErrorID := 0;
   OrderTable[84].OrderNo := 0;
   OrderTable[84].StepNo := 0;
   OrderTable[84].PlaceTime := '';
   OrderTable[84].Device := '';
   OrderTable[84].Sequence := 0;
   OrderTable[84].Status := '';
   OrderTable[84].CompleteTime := '';
   OrderTable[84].ErrorID := 0;
   OrderTable[85].OrderNo := 0;
   OrderTable[85].StepNo := 0;
   OrderTable[85].PlaceTime := '';
   OrderTable[85].Device := '';
   OrderTable[85].Sequence := 0;
   OrderTable[85].Status := '';
   OrderTable[85].CompleteTime := '';
   OrderTable[85].ErrorID := 0;
   OrderTable[86].OrderNo := 0;
   OrderTable[86].StepNo := 0;
   OrderTable[86].PlaceTime := '';
   OrderTable[86].Device := '';
   OrderTable[86].Sequence := 0;
   OrderTable[86].Status := '';
   OrderTable[86].CompleteTime := '';
   OrderTable[86].ErrorID := 0;
   OrderTable[87].OrderNo := 0;
   OrderTable[87].StepNo := 0;
   OrderTable[87].PlaceTime := '';
   OrderTable[87].Device := '';
   OrderTable[87].Sequence := 0;
   OrderTable[87].Status := '';
   OrderTable[87].CompleteTime := '';
   OrderTable[87].ErrorID := 0;
   OrderTable[88].OrderNo := 0;
   OrderTable[88].StepNo := 0;
   OrderTable[88].PlaceTime := '';
   OrderTable[88].Device := '';
   OrderTable[88].Sequence := 0;
   OrderTable[88].Status := '';
   OrderTable[88].CompleteTime := '';
   OrderTable[88].ErrorID := 0;
   OrderTable[89].OrderNo := 0;
   OrderTable[89].StepNo := 0;
   OrderTable[89].PlaceTime := '';
   OrderTable[89].Device := '';
   OrderTable[89].Sequence := 0;
   OrderTable[89].Status := '';
   OrderTable[89].CompleteTime := '';
   OrderTable[89].ErrorID := 0;
   OrderTable[90].OrderNo := 0;
   OrderTable[90].StepNo := 0;
   OrderTable[90].PlaceTime := '';
   OrderTable[90].Device := '';
   OrderTable[90].Sequence := 0;
   OrderTable[90].Status := '';
   OrderTable[90].CompleteTime := '';
   OrderTable[90].ErrorID := 0;
   OrderTable[91].OrderNo := 0;
   OrderTable[91].StepNo := 0;
   OrderTable[91].PlaceTime := '';
   OrderTable[91].Device := '';
   OrderTable[91].Sequence := 0;
   OrderTable[91].Status := '';
   OrderTable[91].CompleteTime := '';
   OrderTable[91].ErrorID := 0;
   OrderTable[92].OrderNo := 0;
   OrderTable[92].StepNo := 0;
   OrderTable[92].PlaceTime := '';
   OrderTable[92].Device := '';
   OrderTable[92].Sequence := 0;
   OrderTable[92].Status := '';
   OrderTable[92].CompleteTime := '';
   OrderTable[92].ErrorID := 0;
   OrderTable[93].OrderNo := 0;
   OrderTable[93].StepNo := 0;
   OrderTable[93].PlaceTime := '';
   OrderTable[93].Device := '';
   OrderTable[93].Sequence := 0;
   OrderTable[93].Status := '';
   OrderTable[93].CompleteTime := '';
   OrderTable[93].ErrorID := 0;
   OrderTable[94].OrderNo := 0;
   OrderTable[94].StepNo := 0;
   OrderTable[94].PlaceTime := '';
   OrderTable[94].Device := '';
   OrderTable[94].Sequence := 0;
   OrderTable[94].Status := '';
   OrderTable[94].CompleteTime := '';
   OrderTable[94].ErrorID := 0;
   OrderTable[95].OrderNo := 0;
   OrderTable[95].StepNo := 0;
   OrderTable[95].PlaceTime := '';
   OrderTable[95].Device := '';
   OrderTable[95].Sequence := 0;
   OrderTable[95].Status := '';
   OrderTable[95].CompleteTime := '';
   OrderTable[95].ErrorID := 0;
   OrderTable[96].OrderNo := 0;
   OrderTable[96].StepNo := 0;
   OrderTable[96].PlaceTime := '';
   OrderTable[96].Device := '';
   OrderTable[96].Sequence := 0;
   OrderTable[96].Status := '';
   OrderTable[96].CompleteTime := '';
   OrderTable[96].ErrorID := 0;
   OrderTable[97].OrderNo := 0;
   OrderTable[97].StepNo := 0;
   OrderTable[97].PlaceTime := '';
   OrderTable[97].Device := '';
   OrderTable[97].Sequence := 0;
   OrderTable[97].Status := '';
   OrderTable[97].CompleteTime := '';
   OrderTable[97].ErrorID := 0;
   OrderTable[98].OrderNo := 0;
   OrderTable[98].StepNo := 0;
   OrderTable[98].PlaceTime := '';
   OrderTable[98].Device := '';
   OrderTable[98].Sequence := 0;
   OrderTable[98].Status := '';
   OrderTable[98].CompleteTime := '';
   OrderTable[98].ErrorID := 0;
   OrderTable[99].OrderNo := 0;
   OrderTable[99].StepNo := 0;
   OrderTable[99].PlaceTime := '';
   OrderTable[99].Device := '';
   OrderTable[99].Sequence := 0;
   OrderTable[99].Status := '';
   OrderTable[99].CompleteTime := '';
   OrderTable[99].ErrorID := 0;
   StepTable[1].OrderNo := 0;
   StepTable[1].StepNo := 0;
   StepTable[1].PlaceTime := '';
   StepTable[1].Device := '';
   StepTable[1].Sequence := 0;
   StepTable[1].Status := '';
   StepTable[1].CompleteTime := '';
   StepTable[1].ErrorID := 0;
   StepTable[2].OrderNo := 0;
   StepTable[2].StepNo := 0;
   StepTable[2].PlaceTime := '';
   StepTable[2].Device := '';
   StepTable[2].Sequence := 0;
   StepTable[2].Status := '';
   StepTable[2].CompleteTime := '';
   StepTable[2].ErrorID := 0;
   StepTable[3].OrderNo := 0;
   StepTable[3].StepNo := 0;
   StepTable[3].PlaceTime := '';
   StepTable[3].Device := '';
   StepTable[3].Sequence := 0;
   StepTable[3].Status := '';
   StepTable[3].CompleteTime := '';
   StepTable[3].ErrorID := 0;
   StepTable[4].OrderNo := 0;
   StepTable[4].StepNo := 0;
   StepTable[4].PlaceTime := '';
   StepTable[4].Device := '';
   StepTable[4].Sequence := 0;
   StepTable[4].Status := '';
   StepTable[4].CompleteTime := '';
   StepTable[4].ErrorID := 0;
   StepTable[5].OrderNo := 0;
   StepTable[5].StepNo := 0;
   StepTable[5].PlaceTime := '';
   StepTable[5].Device := '';
   StepTable[5].Sequence := 0;
   StepTable[5].Status := '';
   StepTable[5].CompleteTime := '';
   StepTable[5].ErrorID := 0;
   StepTable[6].OrderNo := 0;
   StepTable[6].StepNo := 0;
   StepTable[6].PlaceTime := '';
   StepTable[6].Device := '';
   StepTable[6].Sequence := 0;
   StepTable[6].Status := '';
   StepTable[6].CompleteTime := '';
   StepTable[6].ErrorID := 0;
   StepTable[7].OrderNo := 0;
   StepTable[7].StepNo := 0;
   StepTable[7].PlaceTime := '';
   StepTable[7].Device := '';
   StepTable[7].Sequence := 0;
   StepTable[7].Status := '';
   StepTable[7].CompleteTime := '';
   StepTable[7].ErrorID := 0;
   StepTable[8].OrderNo := 0;
   StepTable[8].StepNo := 0;
   StepTable[8].PlaceTime := '';
   StepTable[8].Device := '';
   StepTable[8].Sequence := 0;
   StepTable[8].Status := '';
   StepTable[8].CompleteTime := '';
   StepTable[8].ErrorID := 0;
   StepTable[9].OrderNo := 0;
   StepTable[9].StepNo := 0;
   StepTable[9].PlaceTime := '';
   StepTable[9].Device := '';
   StepTable[9].Sequence := 0;
   StepTable[9].Status := '';
   StepTable[9].CompleteTime := '';
   StepTable[9].ErrorID := 0;
   StepTable[10].OrderNo := 0;
   StepTable[10].StepNo := 0;
   StepTable[10].PlaceTime := '';
   StepTable[10].Device := '';
   StepTable[10].Sequence := 0;
   StepTable[10].Status := '';
   StepTable[10].CompleteTime := '';
   StepTable[10].ErrorID := 0;
   StepTable[11].OrderNo := 0;
   StepTable[11].StepNo := 0;
   StepTable[11].PlaceTime := '';
   StepTable[11].Device := '';
   StepTable[11].Sequence := 0;
   StepTable[11].Status := '';
   StepTable[11].CompleteTime := '';
   StepTable[11].ErrorID := 0;
   StepTable[12].OrderNo := 0;
   StepTable[12].StepNo := 0;
   StepTable[12].PlaceTime := '';
   StepTable[12].Device := '';
   StepTable[12].Sequence := 0;
   StepTable[12].Status := '';
   StepTable[12].CompleteTime := '';
   StepTable[12].ErrorID := 0;
   StepTable[13].OrderNo := 0;
   StepTable[13].StepNo := 0;
   StepTable[13].PlaceTime := '';
   StepTable[13].Device := '';
   StepTable[13].Sequence := 0;
   StepTable[13].Status := '';
   StepTable[13].CompleteTime := '';
   StepTable[13].ErrorID := 0;
   StepTable[14].OrderNo := 0;
   StepTable[14].StepNo := 0;
   StepTable[14].PlaceTime := '';
   StepTable[14].Device := '';
   StepTable[14].Sequence := 0;
   StepTable[14].Status := '';
   StepTable[14].CompleteTime := '';
   StepTable[14].ErrorID := 0;
   StepTable[15].OrderNo := 0;
   StepTable[15].StepNo := 0;
   StepTable[15].PlaceTime := '';
   StepTable[15].Device := '';
   StepTable[15].Sequence := 0;
   StepTable[15].Status := '';
   StepTable[15].CompleteTime := '';
   StepTable[15].ErrorID := 0;
   StepTable[16].OrderNo := 0;
   StepTable[16].StepNo := 0;
   StepTable[16].PlaceTime := '';
   StepTable[16].Device := '';
   StepTable[16].Sequence := 0;
   StepTable[16].Status := '';
   StepTable[16].CompleteTime := '';
   StepTable[16].ErrorID := 0;
   StepTable[17].OrderNo := 0;
   StepTable[17].StepNo := 0;
   StepTable[17].PlaceTime := '';
   StepTable[17].Device := '';
   StepTable[17].Sequence := 0;
   StepTable[17].Status := '';
   StepTable[17].CompleteTime := '';
   StepTable[17].ErrorID := 0;
   StepTable[18].OrderNo := 0;
   StepTable[18].StepNo := 0;
   StepTable[18].PlaceTime := '';
   StepTable[18].Device := '';
   StepTable[18].Sequence := 0;
   StepTable[18].Status := '';
   StepTable[18].CompleteTime := '';
   StepTable[18].ErrorID := 0;
   StepTable[19].OrderNo := 0;
   StepTable[19].StepNo := 0;
   StepTable[19].PlaceTime := '';
   StepTable[19].Device := '';
   StepTable[19].Sequence := 0;
   StepTable[19].Status := '';
   StepTable[19].CompleteTime := '';
   StepTable[19].ErrorID := 0;
   StepTable[20].OrderNo := 0;
   StepTable[20].StepNo := 0;
   StepTable[20].PlaceTime := '';
   StepTable[20].Device := '';
   StepTable[20].Sequence := 0;
   StepTable[20].Status := '';
   StepTable[20].CompleteTime := '';
   StepTable[20].ErrorID := 0;
   CarParked_Confirm := FALSE;
   Running := FALSE;
   IDLE := TRUE;
   Error := FALSE;
   State := 0;
   ResetError := FALSE;
   Ready := TRUE;
   Selected := TRUE;
   Auto_Man := TRUE;
   Paused := FALSE;

END_DATA_BLOCK

DATA_BLOCK "Bypass"
{ S7_Optimized_Access := 'TRUE' }
VERSION : 0.1
NON_RETAIN
   VAR RETAIN
      Main_Panel : "Safety_Bypass_MainPanel";
      Remote_Panel_1 { S7_SetPoint := 'False'} : "Safety_Bypass_RemotePanel";
      Remote_Panel_2 : "Safety_Bypass_RemotePanel";
      Remote_Panel_3 : "Safety_Bypass_RemotePanel";
      Remote_Panel_4 : "Safety_Bypass_RemotePanel";
      Remote_Panel_5 : "Safety_Bypass_RemotePanel";
   END_VAR


BEGIN
   Main_Panel.Estop_Cabinet := FALSE;

END_DATA_BLOCK

DATA_BLOCK "Screen_DB"
{ S7_Optimized_Access := 'TRUE' }
VERSION : 0.1
NON_RETAIN
   VAR
      Settings_ActivePopUp : USInt;
      Alarms_ActiveTable : USInt;
      MainTemplate_ErrorActive : Bool;
      MainTemplate_ErrorCount : USInt;
      MainTemplate_Background : USInt;
      EmptyTemplate_Background : USInt;
      Charge_VTD : Bool;
      Charge_Cnv : Bool;
      Charge_VTD_Commands : Bool;
      Charge_Cnv_Commands : Bool;
      Charge_OT : Bool;
      Shuttle { S7_SetPoint := 'False'} : "Shuttle_MQTT_Status_Msg";
      Shuttle_Select : USInt;
      VTD_Barcode : String;
      VTD_Barcode_Visu : Bool;
      OrderProcessing : Array[1..5] of String;
   END_VAR


BEGIN

END_DATA_BLOCK

DATA_BLOCK "System_DB_2"
{ S7_Optimized_Access := 'TRUE' }
VERSION : 0.1
NON_RETAIN
"System_UDT"

